(* IEC 61131-3 sources: plc-process-lib/tests/POUs/Suites/FB_Valve_Test, 85 files *)

(* ---- ActTimeAccumulatesInRetain.method.decl.st ---- *)
// Время работы привода: 12,5 с с включённым выходом — 12 с в stRetain (доля 0,5 с в накопителе), часы в
// Sts; пока стоит — не копится; шаг времени 60 с идёт в счёт не больше DT_ACCUM_MAX = 10 с. xResetMaint
// обнуляет время «с ТО», полное время не трогает.
METHOD PRIVATE ActTimeAccumulatesInRetain
VAR
    fbTime   : FB_FakeTime;       // подменное время, старт 1 ч
    fbVlv    : FB_Valve;          // арматура под тестом
    stCmd    : ST_ValveCmd;       // команды HMI
    stRetain : ST_DeviceRetain;   // режим Manual по умолчанию, счётчики
    stCfg    : ST_ValveCfg;       // конфигурация (умолчания: Motorized, ZSO и ZSC)
    iStep    : INT;               // шаг цикла
END_VAR

(* ---- ActTimeAccumulatesInRetain.method.impl.st ---- *)
coUnit.TEST('Valve_ActTime_AccumulatesInRetain');

stCfg.tTravel := T#120S;
stRetain.udiOpTime_s := 7190;
fbVlv.xZsc := TRUE;
fbVlv(itfTime := fbTime, stCmd := stCmd, stRetain := stRetain, stCfg := stCfg);
stCmd.xOpen := TRUE;
// t0: выход включён
fbVlv(itfTime := fbTime, stCmd := stCmd, stRetain := stRetain, stCfg := stCfg);
fbVlv.xZsc := FALSE;
FOR iStep := 1 TO 125 DO                                                // 12,5 с
    fbTime.Advance(tStep := T#100MS);
    fbVlv(itfTime := fbTime, stCmd := stCmd, stRetain := stRetain, stCfg := stCfg);
END_FOR
stCmd.xStop := TRUE;
// без шага времени
fbVlv(itfTime := fbTime, stCmd := stCmd, stRetain := stRetain, stCfg := stCfg);
// источник: tools/reference/valve_reference.py, сценарий valve_act_time: 12 с, в накопителе 0,5 с
AssertEquals_UDINT(Expected := 7202, Actual := stRetain.udiOpTime_s, Message := 'total run time 7190 + 12 s');
AssertEquals_UDINT(Expected := 12, Actual := stRetain.udiOpTimeMaint_s, Message := 'run time since maintenance 12 s');
// источник: tools/reference/valve_reference.py, сценарий valve_act_time: hours of 7190 + 12 s
AssertEquals_REAL(Expected := 2.0005555, Actual := fbVlv.stSts.rActTime_h, Delta := 1.0E-6,
                  Message := 'run time in hours');
FOR iStep := 1 TO 20 DO
    fbTime.Advance(tStep := T#100MS);
    fbVlv(itfTime := fbTime, stCmd := stCmd, stRetain := stRetain, stCfg := stCfg);
END_FOR
AssertEquals_UDINT(Expected := 7202, Actual := stRetain.udiOpTime_s, Message := 'no accumulation at rest');
stCmd.xOpen := TRUE;
fbVlv(itfTime := fbTime, stCmd := stCmd, stRetain := stRetain, stCfg := stCfg);
fbTime.Advance(tStep := T#1M);
// один шаг 60 с
fbVlv(itfTime := fbTime, stCmd := stCmd, stRetain := stRetain, stCfg := stCfg);
// источник: tools/reference/valve_reference.py, сценарий valve_act_time: one 60 s step = 10 s (0,5 + 10 с)
AssertEquals_UDINT(Expected := 7212, Actual := stRetain.udiOpTime_s, Message := 'large step bounded by DT_ACCUM_MAX');
stCmd.xResetMaint := TRUE;
fbVlv(itfTime := fbTime, stCmd := stCmd, stRetain := stRetain, stCfg := stCfg);
AssertEquals_UDINT(Expected := 0, Actual := stRetain.udiOpTimeMaint_s,
                   Message := 'xResetMaint clears run time since maintenance');
AssertEquals_UDINT(Expected := 7212, Actual := stRetain.udiOpTime_s, Message := 'total run time kept');

coUnit.TEST_FINISHED();

(* ---- AutoToManualBumpless.method.decl.st ---- *)
// Auto открывает; переход в Manual: цель := текущее направление — ход продолжается до ZSO (арматура не
// дёргается).
METHOD PRIVATE AutoToManualBumpless
VAR
    fbTime   : FB_FakeTime;       // подменное время, старт 1 ч
    fbVlv    : FB_Valve;          // арматура под тестом
    stCmd    : ST_ValveCmd;       // команды HMI
    stRetain : ST_DeviceRetain;   // режим Manual по умолчанию, счётчики
    stCfg    : ST_ValveCfg;       // конфигурация (умолчания: Motorized, ZSO и ZSC)
    iStep    : INT;               // шаг цикла
END_VAR

(* ---- AutoToManualBumpless.method.impl.st ---- *)
coUnit.TEST('Valve_AutoToManual_Bumpless');

stRetain.eRemoteMode := E_DeviceMode.Auto;
fbVlv.xAutoOpen := TRUE;
fbVlv.xZsc := TRUE;
fbVlv(itfTime := fbTime, stCmd := stCmd, stRetain := stRetain, stCfg := stCfg);
AssertTrue(Condition := fbVlv.stSts.eState = E_ValveState.Opening, Message := 'Auto opens on first call');
fbVlv.xZsc := FALSE;
FOR iStep := 1 TO 10 DO
    fbTime.Advance(tStep := T#100MS);
    fbVlv(itfTime := fbTime, stCmd := stCmd, stRetain := stRetain, stCfg := stCfg);
END_FOR
stCmd.stCommon.xSetManual := TRUE;
fbVlv.xAutoOpen := FALSE;
fbTime.Advance(tStep := T#100MS);
fbVlv(itfTime := fbTime, stCmd := stCmd, stRetain := stRetain, stCfg := stCfg);
AssertTrue(Condition := fbVlv.Mode = E_DeviceMode.Manual, Message := 'Manual');
AssertTrue(Condition := fbVlv.stSts.eState = E_ValveState.Opening, Message := 'keeps direction');
AssertTrue(Condition := fbVlv.xQOpen, Message := 'output kept');
FOR iStep := 1 TO 10 DO
    fbTime.Advance(tStep := T#100MS);
    fbVlv.xZso := iStep >= 10;
    fbVlv(itfTime := fbTime, stCmd := stCmd, stRetain := stRetain, stCfg := stCfg);
END_FOR
AssertTrue(Condition := fbVlv.stSts.eState = E_ValveState.Open, Message := 'Open on ZSO');
AssertFalse(Condition := fbVlv.xQOpen, Message := 'output off');

coUnit.TEST_FINISHED();

(* ---- BothLimitsSetsFailureOutputsOff.method.decl.st ---- *)
// Auto, закрыта. Залип ZSO — оба концевика: до tLimitFilter (0,5 с) состояние держится, на 0,5 с —
// BothLimits (wFault бит 2, Failure, тревога слота 2). Запрос автоматики «открыть» выходы не включает,
// Available = FALSE. Отказ не фиксируется: концевик исправен — отказ снят без Reset, Auto ведёт к цели.
METHOD PRIVATE BothLimitsSetsFailureOutputsOff
VAR
    fbTime   : FB_FakeTime;       // подменное время, старт 1 ч
    fbVlv    : FB_Valve;          // арматура под тестом
    stCmd    : ST_ValveCmd;       // команды HMI
    stRetain : ST_DeviceRetain;   // режим Manual по умолчанию, счётчики
    stCfg    : ST_ValveCfg;       // конфигурация (умолчания: Motorized, ZSO и ZSC)
    iStep    : INT;               // шаг цикла
    itfAlm   : I_Alarm;           // слот тревоги через интерфейс
END_VAR

(* ---- BothLimitsSetsFailureOutputsOff.method.impl.st ---- *)
coUnit.TEST('Valve_BothLimits_SetsFailureOutputsOff');

stRetain.eRemoteMode := E_DeviceMode.Auto;
fbVlv.xAutoOpen := FALSE;
fbVlv.xZsc := TRUE;
// Auto, закрыта
fbVlv(itfTime := fbTime, stCmd := stCmd, stRetain := stRetain, stCfg := stCfg);
AssertTrue(Condition := fbVlv.Mode = E_DeviceMode.Auto, Message := 'Auto from retain');
AssertTrue(Condition := fbVlv.stSts.eState = E_ValveState.Closed, Message := 'Closed');
fbVlv.xZso := TRUE;
// t0: оба концевика
fbVlv(itfTime := fbTime, stCmd := stCmd, stRetain := stRetain, stCfg := stCfg);
FOR iStep := 1 TO 4 DO                                                  // t0 + 0,4 с
    fbTime.Advance(tStep := T#100MS);
    fbVlv(itfTime := fbTime, stCmd := stCmd, stRetain := stRetain, stCfg := stCfg);
END_FOR
AssertEquals_WORD(Expected := 0, Actual := fbVlv.stSts.stCommon.wFault, Message := 'no fault before tLimitFilter');
AssertTrue(Condition := fbVlv.stSts.eState = E_ValveState.Closed, Message := 'state held during the filter');
fbTime.Advance(tStep := T#100MS);
// t0 + 0,5 с
fbVlv(itfTime := fbTime, stCmd := stCmd, stRetain := stRetain, stCfg := stCfg);
AssertEquals_WORD(Expected := GVL_Const.VLV_FLT_BOTH_LIMITS, Actual := fbVlv.stSts.stCommon.wFault,
                  Message := 'BothLimits after tLimitFilter');
AssertTrue(Condition := fbVlv.stSts.eState = E_ValveState.Fault, Message := 'Fault state');
AssertTrue(Condition := fbVlv.Status = E_Ne107Status.Failure, Message := 'NE 107 Failure');
itfAlm := fbVlv.GetAlarm(uiIndex := E_ValveAlarm.BothLimits);
AssertTrue(Condition := itfAlm.Active, Message := 'BothLimits alarm active');
fbVlv.xAutoOpen := TRUE;
fbTime.Advance(tStep := T#100MS);
fbVlv(itfTime := fbTime, stCmd := stCmd, stRetain := stRetain, stCfg := stCfg);
AssertFalse(Condition := fbVlv.xQOpen OR fbVlv.xQClose, Message := 'outputs off while both limit switches');
AssertFalse(Condition := fbVlv.Available, Message := 'not available');
fbVlv.xZso := FALSE;
fbTime.Advance(tStep := T#100MS);
// концевик исправен
fbVlv(itfTime := fbTime, stCmd := stCmd, stRetain := stRetain, stCfg := stCfg);
AssertEquals_WORD(Expected := 0, Actual := fbVlv.stSts.stCommon.wFault, Message := 'not latched: clears without Reset');
AssertTrue(Condition := fbVlv.stSts.eState = E_ValveState.Opening, Message := 'Auto resumes towards target');
AssertTrue(Condition := fbVlv.xQOpen, Message := 'open contactor on');

coUnit.TEST_FINISHED();

(* ---- CfgChecksSetBits.method.decl.st ---- *)
// Каждая проверка CheckConfig даёт свой бит wCfgErr: тип вне перечисления; tTravel = 0; Stay у соленоида
// и eSafePos вне перечисления; закрытие по моменту без муфты и муфта у соленоида; tReverse = 0 у
// Motorized (у соленоида допустим); tResetWindow = 0; приоритет тревоги вне перечисления.
METHOD PRIVATE CfgChecksSetBits
VAR
    fbTime   : FB_FakeTime;       // подменное время, старт 1 ч
    fbVlv    : FB_Valve;          // арматура под тестом
    stCmd    : ST_ValveCmd;       // команды HMI
    stRetain : ST_DeviceRetain;   // режим Manual по умолчанию, счётчики
    stCfg    : ST_ValveCfg;       // конфигурация (умолчания: Motorized, ZSO и ZSC)
    uBad     : U_TestValveEnum;   // значения вне строгих перечислений
    stSlot   : ST_AlarmCfg;       // копия слота тревоги
END_VAR

(* ---- CloseLimitReachedGoesClosed.method.decl.st ---- *)
// Manual, задвижка открыта (ZSO). xClose: Closing, включён только xQClose; ZSC на t0 + 3,0 с — Closed,
// выход снят, xClosed. Закрытие циклом «открыто» не считается.
METHOD PRIVATE CloseLimitReachedGoesClosed
VAR
    fbTime   : FB_FakeTime;       // подменное время, старт 1 ч
    fbVlv    : FB_Valve;          // арматура под тестом
    stCmd    : ST_ValveCmd;       // команды HMI
    stRetain : ST_DeviceRetain;   // режим Manual по умолчанию, счётчики
    stCfg    : ST_ValveCfg;       // конфигурация (умолчания: Motorized, ZSO и ZSC)
    iStep    : INT;               // шаг цикла
END_VAR

(* ---- CloseLimitReachedGoesClosed.method.impl.st ---- *)
coUnit.TEST('Valve_Close_LimitReached_GoesClosed');

stCfg.tTravel := T#10S;
fbVlv.xZso := TRUE;
// t0: открыта
fbVlv(itfTime := fbTime, stCmd := stCmd, stRetain := stRetain, stCfg := stCfg);
AssertTrue(Condition := fbVlv.stSts.eState = E_ValveState.Open, Message := 'starts Open on ZSO');
stCmd.xClose := TRUE;
// t0: команда «закрыть»
fbVlv(itfTime := fbTime, stCmd := stCmd, stRetain := stRetain, stCfg := stCfg);
AssertTrue(Condition := fbVlv.stSts.eState = E_ValveState.Closing, Message := 'Closing after xClose');
AssertTrue(Condition := fbVlv.xQClose, Message := 'close contactor on');
AssertFalse(Condition := fbVlv.xQOpen, Message := 'open contactor off');
AssertFalse(Condition := stCmd.xClose, Message := 'xClose cleared');
AssertEquals_WORD(Expected := GVL_Const.VLV_STS_CLOSING,
                  Actual := fbVlv.stSts.stCommon.wStatus AND GVL_Const.VLV_STS_CLOSING, Message := 'CLOSING bit');
FOR iStep := 1 TO 29 DO                                                 // t0 + 0,1 … 2,9 с; ZSO пропал на 0,3 с
    fbTime.Advance(tStep := T#100MS);
    fbVlv.xZso := iStep < 3;
    fbVlv(itfTime := fbTime, stCmd := stCmd, stRetain := stRetain, stCfg := stCfg);
END_FOR
AssertTrue(Condition := fbVlv.xQClose, Message := 'still closing at t0 + 2.9 s');
fbTime.Advance(tStep := T#100MS);
fbVlv.xZsc := TRUE;
// t0 + 3,0 с: ZSC
fbVlv(itfTime := fbTime, stCmd := stCmd, stRetain := stRetain, stCfg := stCfg);
AssertTrue(Condition := fbVlv.stSts.eState = E_ValveState.Closed, Message := 'Closed on ZSC');
AssertFalse(Condition := fbVlv.xQClose, Message := 'contactor off at ZSC');
AssertTrue(Condition := fbVlv.xClosed, Message := 'xClosed');
AssertFalse(Condition := fbVlv.xOpened, Message := 'not xOpened');
AssertEquals_WORD(Expected := GVL_Const.VLV_STS_CLOSED,
                  Actual := fbVlv.stSts.stCommon.wStatus AND (GVL_Const.VLV_STS_OPENED OR GVL_Const.VLV_STS_CLOSED),
                  Message := 'CLOSED bit');
AssertEquals_UDINT(Expected := 0, Actual := stRetain.udiOpCount, Message := 'closing is not an open cycle');

coUnit.TEST_FINISHED();

(* ---- CloseOnTorqueCompletesClosing.method.decl.st ---- *)
// Клиновая задвижка: муфта подключена, закрытие «по моменту». Через 3 с хода сработал ZSC (стоит чуть
// раньше посадки клина) — выход держится; через 0,2 с клин сел, сработала муфта закрытия — Closed без
// отказа, выход снят, xClosed; предупреждения «положение по времени» нет. Муфта отпустила, ZSC держится —
// задвижка остаётся Closed без отказа. Муфта раньше ZSC — тест
// Valve_CloseOnTorque_TorqueBeforeZsc_LatchesTorqueTrip.
METHOD PRIVATE CloseOnTorqueCompletesClosing
VAR
    fbTime   : FB_FakeTime;       // подменное время, старт 1 ч
    fbVlv    : FB_Valve;          // арматура под тестом
    stCmd    : ST_ValveCmd;       // команды HMI
    stRetain : ST_DeviceRetain;   // режим Manual по умолчанию, счётчики
    stCfg    : ST_ValveCfg;       // конфигурация (умолчания: Motorized, ZSO и ZSC)
    iStep    : INT;               // шаг цикла
END_VAR

(* ---- CloseOnTorqueCompletesClosing.method.impl.st ---- *)
coUnit.TEST('Valve_CloseOnTorque_CompletesClosing');

stCfg.xTorqueUsed := TRUE;
stCfg.xCloseOnTorque := TRUE;
fbVlv.xZso := TRUE;
fbVlv(itfTime := fbTime, stCmd := stCmd, stRetain := stRetain, stCfg := stCfg);
stCmd.xClose := TRUE;
fbVlv(itfTime := fbTime, stCmd := stCmd, stRetain := stRetain, stCfg := stCfg);
fbVlv.xZso := FALSE;
FOR iStep := 1 TO 30 DO                                                 // закрывается 3 с
    fbTime.Advance(tStep := T#100MS);
    fbVlv(itfTime := fbTime, stCmd := stCmd, stRetain := stRetain, stCfg := stCfg);
END_FOR
fbVlv.xZsc := TRUE;
FOR iStep := 1 TO 2 DO                                                  // ZSC: клин дожимается 0,2 с
    fbTime.Advance(tStep := T#100MS);
    fbVlv(itfTime := fbTime, stCmd := stCmd, stRetain := stRetain, stCfg := stCfg);
END_FOR
AssertTrue(Condition := fbVlv.xQClose, Message := 'output held on ZSC until torque');
fbVlv.xTorqueClose := TRUE;
fbTime.Advance(tStep := T#100MS);
// клин сел: муфта закрытия
fbVlv(itfTime := fbTime, stCmd := stCmd, stRetain := stRetain, stCfg := stCfg);
AssertTrue(Condition := fbVlv.stSts.eState = E_ValveState.Closed, Message := 'Closed on torque');
AssertFalse(Condition := fbVlv.xQClose, Message := 'output off');
AssertEquals_WORD(Expected := 0, Actual := fbVlv.stSts.stCommon.wFault, Message := 'no torque trip');
AssertTrue(Condition := fbVlv.xClosed, Message := 'xClosed');
AssertEquals_WORD(Expected := 0, Actual := fbVlv.stSts.stCommon.wWarning AND GVL_Const.VLV_WRN_POSITION_BY_TIME,
                  Message := 'closed by torque, not by time');
fbVlv.xTorqueClose := FALSE;
FOR iStep := 1 TO 20 DO                                                 // 2 с: муфта отпустила, ZSC держится
    fbTime.Advance(tStep := T#100MS);
    fbVlv(itfTime := fbTime, stCmd := stCmd, stRetain := stRetain, stCfg := stCfg);
END_FOR
AssertEquals_WORD(Expected := 0, Actual := fbVlv.stSts.stCommon.wFault, Message := 'no fault after torque released');
AssertTrue(Condition := fbVlv.stSts.eState = E_ValveState.Closed, Message := 'stays Closed');

coUnit.TEST_FINISHED();

(* ---- CloseOnTorqueNoZscTorqueMissingSetsFailToClose.method.decl.st ---- *)
// Клиновая задвижка без ZSC (xZscUsed = FALSE), закрытие «по моменту», tTravel = 10 с. Муфта закрытия
// так и не сработала: на t0 + 9,9 с ещё Closing и выход «закрывать» держится, ровно на t0 + 10,0 с —
// FailToClose, выход снят, xClosed нет. Положения «закрыто по времени» у закрытия по моменту нет: его
// подтверждает только муфта.
METHOD PRIVATE CloseOnTorqueNoZscTorqueMissingSetsFailToClose
VAR
    fbTime   : FB_FakeTime;       // подменное время, старт 1 ч
    fbVlv    : FB_Valve;          // арматура под тестом
    stCmd    : ST_ValveCmd;       // команды HMI
    stRetain : ST_DeviceRetain;   // режим Manual по умолчанию, счётчики
    stCfg    : ST_ValveCfg;       // конфигурация: без ZSC, закрытие по моменту
    iStep    : INT;               // шаг цикла
END_VAR

(* ---- CloseOnTorqueNoZscTorqueMissingSetsFailToClose.method.impl.st ---- *)
coUnit.TEST('Valve_CloseOnTorqueNoZsc_TorqueMissing_SetsFailToClose');

stCfg.xZscUsed := FALSE;
stCfg.xTorqueUsed := TRUE;
stCfg.xCloseOnTorque := TRUE;
stCfg.tTravel := T#10S;
fbVlv.xZso := TRUE;
fbVlv(itfTime := fbTime, stCmd := stCmd, stRetain := stRetain, stCfg := stCfg);
stCmd.xClose := TRUE;
// t0: Closing
fbVlv(itfTime := fbTime, stCmd := stCmd, stRetain := stRetain, stCfg := stCfg);
fbVlv.xZso := FALSE;
FOR iStep := 1 TO 99 DO                                                 // до t0 + 9,9 с, муфты нет
    fbTime.Advance(tStep := T#100MS);
    fbVlv(itfTime := fbTime, stCmd := stCmd, stRetain := stRetain, stCfg := stCfg);
END_FOR
AssertTrue(Condition := fbVlv.stSts.eState = E_ValveState.Closing, Message := 'still closing at t0 + 9.9 s');
AssertTrue(Condition := fbVlv.xQClose, Message := 'close output held until torque');
fbTime.Advance(tStep := T#100MS);
// t0 + 10,0 с
fbVlv(itfTime := fbTime, stCmd := stCmd, stRetain := stRetain, stCfg := stCfg);
AssertTrue(Condition := fbVlv.stSts.eState = E_ValveState.Fault, Message := 'Fault at tTravel, not closed by time');
AssertEquals_WORD(Expected := GVL_Const.VLV_FLT_FAIL_TO_CLOSE, Actual := fbVlv.stSts.stCommon.wFault,
                  Message := 'wFault FailToClose');
AssertFalse(Condition := fbVlv.xQClose, Message := 'output off on timeout');
AssertFalse(Condition := fbVlv.xClosed, Message := 'not reported closed');

coUnit.TEST_FINISHED();

(* ---- CloseOnTorqueTorqueBeforeZscLatchesTorqueTrip.method.decl.st ---- *)
// Клиновая задвижка, закрытие «по моменту», ZSC подключён. Муфта закрытия сработала на t0 + 3 с, а
// ZSC — нет: ZSC настроен чуть раньше посадки клина (VLV-19), значит, это не посадка, а заклинивание или
// посторонний предмет — TorqueTrip, выход снят, xClosed нет. Тот же ход без ZSC (xZscUsed = FALSE):
// муфта — штатное окончание закрытия, Closed без отказа, и после того как муфта отпустила, задвижка
// остаётся Closed.
METHOD PRIVATE CloseOnTorqueTorqueBeforeZscLatchesTorqueTrip
VAR
    fbTime    : FB_FakeTime;       // подменное время, старт 1 ч
    fbVlv     : FB_Valve;          // задвижка с ZSC
    stCmd     : ST_ValveCmd;       // команды HMI
    stRetain  : ST_DeviceRetain;   // режим Manual по умолчанию, счётчики
    stCfg     : ST_ValveCfg;       // конфигурация (умолчания: Motorized, ZSO и ZSC)
    fbVlv2    : FB_Valve;          // задвижка без ZSC
    stCmd2    : ST_ValveCmd;       // команды HMI второй задвижки
    stRetain2 : ST_DeviceRetain;   // режим Manual по умолчанию
    stCfg2    : ST_ValveCfg;       // конфигурация второй задвижки
    iStep     : INT;               // шаг цикла
END_VAR

(* ---- CloseOnTorqueTorqueBeforeZscLatchesTorqueTrip.method.impl.st ---- *)
coUnit.TEST('Valve_CloseOnTorque_TorqueBeforeZsc_LatchesTorqueTrip');

stCfg.xTorqueUsed := TRUE;
stCfg.xCloseOnTorque := TRUE;
fbVlv.xZso := TRUE;
fbVlv(itfTime := fbTime, stCmd := stCmd, stRetain := stRetain, stCfg := stCfg);
stCmd.xClose := TRUE;
fbVlv(itfTime := fbTime, stCmd := stCmd, stRetain := stRetain, stCfg := stCfg);
fbVlv.xZso := FALSE;
FOR iStep := 1 TO 30 DO                                                 // закрывается 3 с
    fbTime.Advance(tStep := T#100MS);
    fbVlv(itfTime := fbTime, stCmd := stCmd, stRetain := stRetain, stCfg := stCfg);
END_FOR
fbVlv.xTorqueClose := TRUE;
fbTime.Advance(tStep := T#100MS);
// муфта раньше ZSC
fbVlv(itfTime := fbTime, stCmd := stCmd, stRetain := stRetain, stCfg := stCfg);
AssertTrue(Condition := fbVlv.stSts.eState = E_ValveState.Fault, Message := 'torque before ZSC: Fault');
AssertEquals_WORD(Expected := GVL_Const.VLV_FLT_TORQUE_TRIP, Actual := fbVlv.stSts.stCommon.wFault,
                  Message := 'wFault TorqueTrip');
AssertFalse(Condition := fbVlv.xQClose, Message := 'output off');
AssertFalse(Condition := fbVlv.xClosed, Message := 'not reported closed');

stCfg2.xZscUsed := FALSE;
stCfg2.xTorqueUsed := TRUE;
stCfg2.xCloseOnTorque := TRUE;
fbVlv2.xZso := TRUE;
fbVlv2(itfTime := fbTime, stCmd := stCmd2, stRetain := stRetain2, stCfg := stCfg2);
stCmd2.xClose := TRUE;
fbVlv2(itfTime := fbTime, stCmd := stCmd2, stRetain := stRetain2, stCfg := stCfg2);
fbVlv2.xZso := FALSE;
FOR iStep := 1 TO 30 DO                                                 // закрывается 3 с
    fbTime.Advance(tStep := T#100MS);
    fbVlv2(itfTime := fbTime, stCmd := stCmd2, stRetain := stRetain2, stCfg := stCfg2);
END_FOR
fbVlv2.xTorqueClose := TRUE;
fbTime.Advance(tStep := T#100MS);
// без ZSC муфта — окончание закрытия
fbVlv2(itfTime := fbTime, stCmd := stCmd2, stRetain := stRetain2, stCfg := stCfg2);
AssertTrue(Condition := fbVlv2.stSts.eState = E_ValveState.Closed, Message := 'no ZSC: Closed on torque');
AssertEquals_WORD(Expected := 0, Actual := fbVlv2.stSts.stCommon.wFault, Message := 'no ZSC: no torque trip');
AssertFalse(Condition := fbVlv2.xQClose, Message := 'no ZSC: output off');
AssertTrue(Condition := fbVlv2.xClosed, Message := 'no ZSC: xClosed');
fbVlv2.xTorqueClose := FALSE;
FOR iStep := 1 TO 20 DO                                                 // муфта отпустила, 2 с
    fbTime.Advance(tStep := T#100MS);
    fbVlv2(itfTime := fbTime, stCmd := stCmd2, stRetain := stRetain2, stCfg := stCfg2);
END_FOR
AssertTrue(Condition := fbVlv2.stSts.eState = E_ValveState.Closed, Message := 'no ZSC: stays Closed');
AssertEquals_WORD(Expected := 0, Actual := fbVlv2.stSts.stCommon.wFault, Message := 'no ZSC: still no fault');

coUnit.TEST_FINISHED();

(* ---- CloseOnTorqueZscAloneKeepsDrivingUntilTimeout.method.decl.st ---- *)
// Клиновая задвижка, закрытие «по моменту», tTravel = 10 с. ZSC сработал на t0 + 3 с (концевик стоит
// чуть раньше посадки клина): выход «закрывать» не снимается — клин дожимается до муфты, xClosed нет.
// Муфта так и не сработала: ровно на t0 + 10,0 с — FailToClose, выход снят; положение по ZSC видно в
// xClosed. Reset снимает отказ — далее состояние по концевикам (Closed).
METHOD PRIVATE CloseOnTorqueZscAloneKeepsDrivingUntilTimeout
VAR
    fbTime   : FB_FakeTime;       // подменное время, старт 1 ч
    fbVlv    : FB_Valve;          // арматура под тестом
    stCmd    : ST_ValveCmd;       // команды HMI
    stRetain : ST_DeviceRetain;   // режим Manual по умолчанию, счётчики
    stCfg    : ST_ValveCfg;       // конфигурация (умолчания: Motorized, ZSO и ZSC)
    iStep    : INT;               // шаг цикла
END_VAR

(* ---- CloseOnTorqueZscAloneKeepsDrivingUntilTimeout.method.impl.st ---- *)
coUnit.TEST('Valve_CloseOnTorque_ZscAloneKeepsDrivingUntilTimeout');

stCfg.tTravel := T#10S;
stCfg.xTorqueUsed := TRUE;
stCfg.xCloseOnTorque := TRUE;
fbVlv.xZso := TRUE;
// t0: открыта
fbVlv(itfTime := fbTime, stCmd := stCmd, stRetain := stRetain, stCfg := stCfg);
stCmd.xClose := TRUE;
// t0: Closing
fbVlv(itfTime := fbTime, stCmd := stCmd, stRetain := stRetain, stCfg := stCfg);
fbVlv.xZso := FALSE;
FOR iStep := 1 TO 30 DO                                                 // до t0 + 3,0 с
    fbTime.Advance(tStep := T#100MS);
    fbVlv(itfTime := fbTime, stCmd := stCmd, stRetain := stRetain, stCfg := stCfg);
END_FOR
fbVlv.xZsc := TRUE;
FOR iStep := 1 TO 69 DO                                                 // ZSC есть, муфты нет: до t0 + 9,9 с
    fbTime.Advance(tStep := T#100MS);
    fbVlv(itfTime := fbTime, stCmd := stCmd, stRetain := stRetain, stCfg := stCfg);
END_FOR
AssertTrue(Condition := fbVlv.stSts.eState = E_ValveState.Closing, Message := 'still closing on ZSC alone');
AssertTrue(Condition := fbVlv.xQClose, Message := 'close output held until torque');
AssertFalse(Condition := fbVlv.xClosed, Message := 'not closed before torque');
AssertEquals_WORD(Expected := 0, Actual := fbVlv.stSts.stCommon.wFault, Message := 'no fault before tTravel');
fbTime.Advance(tStep := T#100MS);
// t0 + 10,0 с: муфта не сработала
fbVlv(itfTime := fbTime, stCmd := stCmd, stRetain := stRetain, stCfg := stCfg);
AssertTrue(Condition := fbVlv.stSts.eState = E_ValveState.Fault, Message := 'Fault at tTravel');
AssertEquals_WORD(Expected := GVL_Const.VLV_FLT_FAIL_TO_CLOSE, Actual := fbVlv.stSts.stCommon.wFault,
                  Message := 'wFault FailToClose');
AssertFalse(Condition := fbVlv.xQClose, Message := 'output off on timeout');
AssertTrue(Condition := fbVlv.xClosed, Message := 'ZSC position visible in Fault');
stCmd.stCommon.xReset := TRUE;
fbVlv(itfTime := fbTime, stCmd := stCmd, stRetain := stRetain, stCfg := stCfg);
AssertEquals_WORD(Expected := 0, Actual := fbVlv.stSts.stCommon.wFault, Message := 'cleared by Reset');
AssertTrue(Condition := fbVlv.stSts.eState = E_ValveState.Closed, Message := 'Closed by ZSC after Reset');
AssertFalse(Condition := fbVlv.xQClose, Message := 'no output after Reset');

coUnit.TEST_FINISHED();

(* ---- CyclesCountedOnOpen.method.decl.st ---- *)
// Цикл — вход в Open, если прошлое крайнее положение не Open: открыть (1), закрыть (1), открыть (2) —
// stRetain и stSts. Неполный ход Open -> стоп -> снова Open циклом не считается. xResetMaint обнуляет
// счётчик «с ТО», полный не трогает. Перед каждой сменой направления арматура стоит 1 с: встречный ход
// начинается не раньше tReverse после снятия выхода (тест Valve_ReverseAfterEndStop_WaitsReversePause).
METHOD PRIVATE CyclesCountedOnOpen
VAR
    fbTime   : FB_FakeTime;       // подменное время, старт 1 ч
    fbVlv    : FB_Valve;          // арматура под тестом
    stCmd    : ST_ValveCmd;       // команды HMI
    stRetain : ST_DeviceRetain;   // режим Manual по умолчанию, счётчики
    stCfg    : ST_ValveCfg;       // конфигурация (умолчания: Motorized, ZSO и ZSC)
    iStep    : INT;               // шаг цикла
END_VAR

(* ---- CyclesCountedOnOpen.method.impl.st ---- *)
coUnit.TEST('Valve_Cycles_CountedOnOpen');

fbVlv.xZsc := TRUE;
fbVlv(itfTime := fbTime, stCmd := stCmd, stRetain := stRetain, stCfg := stCfg);
stCmd.xOpen := TRUE;
fbVlv(itfTime := fbTime, stCmd := stCmd, stRetain := stRetain, stCfg := stCfg);
FOR iStep := 1 TO 10 DO
    fbTime.Advance(tStep := T#100MS);
    fbVlv.xZsc := FALSE;
    fbVlv.xZso := iStep >= 10;
    fbVlv(itfTime := fbTime, stCmd := stCmd, stRetain := stRetain, stCfg := stCfg);
END_FOR
AssertEquals_UDINT(Expected := 1, Actual := stRetain.udiOpCount, Message := 'first open: 1');
FOR iStep := 1 TO 10 DO                                                 // стоит 1 с (выбег, tReverse)
    fbTime.Advance(tStep := T#100MS);
    fbVlv(itfTime := fbTime, stCmd := stCmd, stRetain := stRetain, stCfg := stCfg);
END_FOR
stCmd.xClose := TRUE;
fbVlv(itfTime := fbTime, stCmd := stCmd, stRetain := stRetain, stCfg := stCfg);
FOR iStep := 1 TO 10 DO
    fbTime.Advance(tStep := T#100MS);
    fbVlv.xZso := FALSE;
    fbVlv.xZsc := iStep >= 10;
    fbVlv(itfTime := fbTime, stCmd := stCmd, stRetain := stRetain, stCfg := stCfg);
END_FOR
AssertTrue(Condition := fbVlv.stSts.eState = E_ValveState.Closed, Message := 'Closed');
AssertEquals_UDINT(Expected := 1, Actual := stRetain.udiOpCount, Message := 'closing does not count');
FOR iStep := 1 TO 10 DO                                                 // стоит 1 с (выбег, tReverse)
    fbTime.Advance(tStep := T#100MS);
    fbVlv(itfTime := fbTime, stCmd := stCmd, stRetain := stRetain, stCfg := stCfg);
END_FOR
stCmd.xOpen := TRUE;
fbVlv(itfTime := fbTime, stCmd := stCmd, stRetain := stRetain, stCfg := stCfg);
FOR iStep := 1 TO 10 DO
    fbTime.Advance(tStep := T#100MS);
    fbVlv.xZsc := FALSE;
    fbVlv.xZso := iStep >= 10;
    fbVlv(itfTime := fbTime, stCmd := stCmd, stRetain := stRetain, stCfg := stCfg);
END_FOR
AssertEquals_UDINT(Expected := 2, Actual := stRetain.udiOpCount, Message := 'second open: 2');
AssertEquals_UDINT(Expected := 2, Actual := stRetain.udiOpCountMaint, Message := 'maintenance counter 2');
AssertEquals_UDINT(Expected := 2, Actual := fbVlv.stSts.udiCycles, Message := 'Sts udiCycles');
AssertEquals_UDINT(Expected := 2, Actual := fbVlv.stSts.udiCyclesMaint, Message := 'Sts udiCyclesMaint');
FOR iStep := 1 TO 10 DO                                                 // стоит 1 с (выбег, tReverse)
    fbTime.Advance(tStep := T#100MS);
    fbVlv(itfTime := fbTime, stCmd := stCmd, stRetain := stRetain, stCfg := stCfg);
END_FOR
stCmd.xClose := TRUE;
fbVlv(itfTime := fbTime, stCmd := stCmd, stRetain := stRetain, stCfg := stCfg);
FOR iStep := 1 TO 5 DO
    fbTime.Advance(tStep := T#100MS);
    fbVlv.xZso := FALSE;
    fbVlv(itfTime := fbTime, stCmd := stCmd, stRetain := stRetain, stCfg := stCfg);
END_FOR
stCmd.xStop := TRUE;
fbVlv(itfTime := fbTime, stCmd := stCmd, stRetain := stRetain, stCfg := stCfg);
FOR iStep := 1 TO 10 DO                                                 // стоит 1 с (выбег, tReverse)
    fbTime.Advance(tStep := T#100MS);
    fbVlv(itfTime := fbTime, stCmd := stCmd, stRetain := stRetain, stCfg := stCfg);
END_FOR
stCmd.xOpen := TRUE;
fbVlv(itfTime := fbTime, stCmd := stCmd, stRetain := stRetain, stCfg := stCfg);
FOR iStep := 1 TO 5 DO
    fbTime.Advance(tStep := T#100MS);
    fbVlv.xZso := iStep >= 5;
    fbVlv(itfTime := fbTime, stCmd := stCmd, stRetain := stRetain, stCfg := stCfg);
END_FOR
AssertTrue(Condition := fbVlv.stSts.eState = E_ValveState.Open, Message := 'Open again');
AssertEquals_UDINT(Expected := 2, Actual := stRetain.udiOpCount,
                   Message := 'partial stroke back to Open is not a cycle');
stCmd.xResetMaint := TRUE;
fbVlv(itfTime := fbTime, stCmd := stCmd, stRetain := stRetain, stCfg := stCfg);
AssertEquals_UDINT(Expected := 0, Actual := stRetain.udiOpCountMaint, Message := 'maintenance counter reset');
AssertEquals_UDINT(Expected := 2, Actual := stRetain.udiOpCount, Message := 'total kept');
AssertTrue(Condition := fbVlv.stSts.stCommon.eCmdResult = E_CmdResult.Accepted, Message := 'xResetMaint accepted');
AssertFalse(Condition := stCmd.xResetMaint, Message := 'xResetMaint cleared');

coUnit.TEST_FINISHED();

(* ---- DefaultCfgPassesCheck.method.decl.st ---- *)
// Умолчания ST_ValveCfg проходят CheckConfig; тип в stCommon — Valve, слотов тревог 7; приоритеты по
// умолчанию (FailToOpen — Medium, InterlockAct — None); слот 7 не используется; NE 107 Good.
METHOD PRIVATE DefaultCfgPassesCheck
VAR
    fbTime   : FB_FakeTime;       // подменное время, старт 1 ч
    fbVlv    : FB_Valve;          // арматура под тестом
    stCmd    : ST_ValveCmd;       // команды HMI
    stRetain : ST_DeviceRetain;   // режим Manual по умолчанию, счётчики
    stCfg    : ST_ValveCfg;       // конфигурация (умолчания: Motorized, ZSO и ZSC)
    itfAlm   : I_Alarm;           // слот тревоги через интерфейс
END_VAR

(* ---- ExtFaultTripsAndResetRejectedWhileActive.method.decl.st ---- *)
// Внешняя авария в ходе: Fault, выход снят, тревога слота 5 с номером udiAlarmIdBase + 5. Reset при
// действующей причине: Accepted сразу, окно tResetWindow = 3 с; до конца окна второго результата нет,
// ровно на 3 с — RejectedFault, отказ остаётся. Причина ушла — отказ держится до Reset; Reset снимает.
METHOD PRIVATE ExtFaultTripsAndResetRejectedWhileActive
VAR
    fbTime   : FB_FakeTime;       // подменное время, старт 1 ч
    fbVlv    : FB_Valve;          // арматура под тестом
    stCmd    : ST_ValveCmd;       // команды HMI
    stRetain : ST_DeviceRetain;   // режим Manual по умолчанию, счётчики
    stCfg    : ST_ValveCfg;       // конфигурация (умолчания: Motorized, ZSO и ZSC)
    iStep    : INT;               // шаг цикла
    itfAlm   : I_Alarm;           // слот тревоги через интерфейс
    uiSeq    : UINT;              // номер команды до Reset
END_VAR

(* ---- ExtFaultTripsAndResetRejectedWhileActive.method.impl.st ---- *)
coUnit.TEST('Valve_ExtFault_TripsAndResetRejectedWhileActive');

stCfg.udiAlarmIdBase := 120;
fbVlv.xZsc := TRUE;
fbVlv(itfTime := fbTime, stCmd := stCmd, stRetain := stRetain, stCfg := stCfg);
stCmd.xOpen := TRUE;
fbVlv(itfTime := fbTime, stCmd := stCmd, stRetain := stRetain, stCfg := stCfg);
fbVlv.xZsc := FALSE;
fbTime.Advance(tStep := T#100MS);
fbVlv(itfTime := fbTime, stCmd := stCmd, stRetain := stRetain, stCfg := stCfg);
fbVlv.xExtFault := TRUE;
fbTime.Advance(tStep := T#100MS);
fbVlv(itfTime := fbTime, stCmd := stCmd, stRetain := stRetain, stCfg := stCfg);
AssertTrue(Condition := fbVlv.stSts.eState = E_ValveState.Fault, Message := 'Fault on external fault');
AssertFalse(Condition := fbVlv.xQOpen, Message := 'output off');
AssertEquals_WORD(Expected := GVL_Const.VLV_FLT_EXT_FAULT, Actual := fbVlv.stSts.stCommon.wFault,
                  Message := 'wFault ExtFault');
itfAlm := fbVlv.GetAlarm(uiIndex := E_ValveAlarm.ExtFault);
AssertEquals_UDINT(Expected := 125, Actual := itfAlm.Id, Message := 'alarm id = base + slot');
AssertTrue(Condition := itfAlm.State = E_AlarmState.ActiveUnack, Message := 'ExtFault alarm');
uiSeq := fbVlv.stSts.stCommon.uiCmdSeq;
stCmd.stCommon.xReset := TRUE;
// t1: Reset, причина действует
fbVlv(itfTime := fbTime, stCmd := stCmd, stRetain := stRetain, stCfg := stCfg);
AssertTrue(Condition := fbVlv.stSts.stCommon.eCmdResult = E_CmdResult.Accepted, Message := 'Reset accepted');
AssertEquals_UINT(Expected := uiSeq + 1, Actual := fbVlv.stSts.stCommon.uiCmdSeq, Message := 'one result so far');
FOR iStep := 1 TO 29 DO                                                 // t1 + 2,9 с
    fbTime.Advance(tStep := T#100MS);
    fbVlv(itfTime := fbTime, stCmd := stCmd, stRetain := stRetain, stCfg := stCfg);
END_FOR
AssertEquals_UINT(Expected := uiSeq + 1, Actual := fbVlv.stSts.stCommon.uiCmdSeq,
                  Message := 'no second result before the window ends');
fbTime.Advance(tStep := T#100MS);
// t1 + 3,0 с
fbVlv(itfTime := fbTime, stCmd := stCmd, stRetain := stRetain, stCfg := stCfg);
AssertTrue(Condition := fbVlv.stSts.stCommon.eCmdResult = E_CmdResult.RejectedFault,
           Message := 'RejectedFault at the window end');
AssertEquals_UINT(Expected := uiSeq + 2, Actual := fbVlv.stSts.stCommon.uiCmdSeq, Message := 'second result');
AssertEquals_WORD(Expected := GVL_Const.VLV_FLT_EXT_FAULT, Actual := fbVlv.stSts.stCommon.wFault,
                  Message := 'still faulted');
fbVlv.xExtFault := FALSE;
fbTime.Advance(tStep := T#100MS);
fbVlv(itfTime := fbTime, stCmd := stCmd, stRetain := stRetain, stCfg := stCfg);
AssertEquals_WORD(Expected := GVL_Const.VLV_FLT_EXT_FAULT, Actual := fbVlv.stSts.stCommon.wFault,
                  Message := 'latched after the cause is gone');
stCmd.stCommon.xReset := TRUE;
fbVlv(itfTime := fbTime, stCmd := stCmd, stRetain := stRetain, stCfg := stCfg);
AssertEquals_WORD(Expected := 0, Actual := fbVlv.stSts.stCommon.wFault, Message := 'cleared by Reset');
AssertTrue(Condition := fbVlv.stSts.stCommon.eCmdResult = E_CmdResult.Accepted, Message := 'Reset accepted');
fbTime.Advance(tStep := T#100MS);
fbVlv(itfTime := fbTime, stCmd := stCmd, stRetain := stRetain, stCfg := stCfg);
AssertTrue(Condition := itfAlm.State = E_AlarmState.Normal, Message := 'alarm Normal after Reset');
AssertTrue(Condition := fbVlv.stSts.eState = E_ValveState.Intermediate, Message := 'Intermediate');

coUnit.TEST_FINISHED();

(* ---- InterlockAfterPositionLostDrivesSafe.method.decl.st ---- *)
// Задвижка в Auto открыта по ZSO; ZSO пропал (обрыв) — через tLimitFilter зафиксирован PositionLost, выходов нет.
// Блокировка (Closed): задвижка закрывается (VLV-20); ход заканчивается по ZSC — он согласован (ZSO нет). Отказ
// держится до Reset; после Reset — Closed по концевикам, движения нет (уже в положении безопасности).
METHOD PRIVATE InterlockAfterPositionLostDrivesSafe
VAR
    fbTime   : FB_FakeTime;       // подменное время, старт 1 ч
    fbVlv    : FB_Valve;          // арматура под тестом
    stCmd    : ST_ValveCmd;       // команды HMI
    stRetain : ST_DeviceRetain;   // режим, счётчики
    stCfg    : ST_ValveCfg;       // конфигурация (умолчания: Motorized, ZSO и ZSC)
    iStep    : INT;               // шаг цикла
END_VAR

(* ---- InterlockAfterPositionLostDrivesSafe.method.impl.st ---- *)
coUnit.TEST('Valve_InterlockAfterPositionLost_DrivesSafe');

stRetain.eRemoteMode := E_DeviceMode.Auto;
fbVlv.xAutoOpen := TRUE;
fbVlv.xZso := TRUE;
fbVlv(itfTime := fbTime, stCmd := stCmd, stRetain := stRetain, stCfg := stCfg);       // t0: Open по ZSO
fbVlv.xZso := FALSE;                                                                   // обрыв ZSO
FOR iStep := 1 TO 6 DO                                                               // фильтр 0,5 с
    fbTime.Advance(tStep := T#100MS);
    fbVlv(itfTime := fbTime, stCmd := stCmd, stRetain := stRetain, stCfg := stCfg);
END_FOR
AssertEquals_WORD(Expected := GVL_Const.VLV_FLT_POSITION_LOST, Actual := fbVlv.stSts.stCommon.wFault,
                  Message := 'precondition: PositionLost latched');
AssertFalse(Condition := fbVlv.xQOpen OR fbVlv.xQClose, Message := 'no motion with the fault alone');
fbVlv.wInterlock := 16#0001;
fbTime.Advance(tStep := T#100MS);
fbVlv(itfTime := fbTime, stCmd := stCmd, stRetain := stRetain, stCfg := stCfg);       // t1: блокировка
AssertTrue(Condition := fbVlv.xQClose, Message := 'interlock drives Closed despite PositionLost');
FOR iStep := 1 TO 30 DO
    fbTime.Advance(tStep := T#100MS);
    fbVlv(itfTime := fbTime, stCmd := stCmd, stRetain := stRetain, stCfg := stCfg);
END_FOR
AssertTrue(Condition := fbVlv.xQClose, Message := 'still closing before ZSC');
fbVlv.xZsc := TRUE;
fbTime.Advance(tStep := T#100MS);
fbVlv(itfTime := fbTime, stCmd := stCmd, stRetain := stRetain, stCfg := stCfg);       // ZSC
AssertFalse(Condition := fbVlv.xQClose, Message := 'safe move ends on a consistent ZSC');
AssertTrue(Condition := fbVlv.xClosed, Message := 'position Closed shown');
AssertEquals_WORD(Expected := GVL_Const.VLV_FLT_POSITION_LOST, Actual := fbVlv.stSts.stCommon.wFault,
                  Message := 'fault latched until Reset');
stCmd.stCommon.xReset := TRUE;
fbTime.Advance(tStep := T#100MS);
fbVlv(itfTime := fbTime, stCmd := stCmd, stRetain := stRetain, stCfg := stCfg);
AssertEquals_WORD(Expected := 0, Actual := fbVlv.stSts.stCommon.wFault, Message := 'cleared by Reset');
AssertTrue(Condition := fbVlv.stSts.eState = E_ValveState.Closed, Message := 'Closed after Reset');
AssertFalse(Condition := fbVlv.xQOpen OR fbVlv.xQClose, Message := 'no motion: already in the safe position');

coUnit.TEST_FINISHED();

(* ---- InterlockDrivesToSafePosition.method.decl.st ---- *)
// Manual, открыта, разрешения на закрытие нет (xClose — RejectedPermit). Блокировка (биты 3 и 4) ведёт в
// положение безопасности Closed без разрешения: Closing, бит INTERLOCKED, wInterlock, первопричина —
// младший бит 3. Команды — RejectedInterlock; новый бит первопричину не меняет. После снятия блокировки
// Manual остаётся закрытым; первопричина держится до Reset.
METHOD PRIVATE InterlockDrivesToSafePosition
VAR
    fbTime   : FB_FakeTime;       // подменное время, старт 1 ч
    fbVlv    : FB_Valve;          // арматура под тестом
    stCmd    : ST_ValveCmd;       // команды HMI
    stRetain : ST_DeviceRetain;   // режим Manual по умолчанию, счётчики
    stCfg    : ST_ValveCfg;       // конфигурация (умолчания: Motorized, ZSO и ZSC)
    iStep    : INT;               // шаг цикла
END_VAR

(* ---- InterlockDrivesToSafePosition.method.impl.st ---- *)
coUnit.TEST('Valve_Interlock_DrivesToSafePosition');

fbVlv.xZso := TRUE;
fbVlv.wPermitClose := 16#0000;
// открыта, закрывать нельзя
fbVlv(itfTime := fbTime, stCmd := stCmd, stRetain := stRetain, stCfg := stCfg);
stCmd.xClose := TRUE;
fbVlv(itfTime := fbTime, stCmd := stCmd, stRetain := stRetain, stCfg := stCfg);
AssertTrue(Condition := fbVlv.stSts.stCommon.eCmdResult = E_CmdResult.RejectedPermit,
           Message := 'close without permit rejected');
AssertTrue(Condition := fbVlv.stSts.eState = E_ValveState.Open, Message := 'still Open');
fbVlv.wInterlock := 16#0018;
fbTime.Advance(tStep := T#100MS);
// блокировка
fbVlv(itfTime := fbTime, stCmd := stCmd, stRetain := stRetain, stCfg := stCfg);
AssertTrue(Condition := fbVlv.stSts.eState = E_ValveState.Closing, Message := 'interlock drives Closed');
AssertTrue(Condition := fbVlv.xQClose, Message := 'close contactor on without permit');
AssertEquals_WORD(Expected := GVL_Const.VLV_STS_INTERLOCKED,
                  Actual := fbVlv.stSts.stCommon.wStatus AND GVL_Const.VLV_STS_INTERLOCKED,
Message := 'INTERLOCKED bit');
AssertEquals_WORD(Expected := 16#0018, Actual := fbVlv.stSts.wInterlock, Message := 'active interlocks');
AssertEquals_UINT(Expected := 3, Actual := fbVlv.stSts.uiFirstOut, Message := 'first out = lowest new bit');
AssertEquals_WORD(Expected := 0, Actual := fbVlv.stSts.wPermitMissing, Message := 'no permit needed');
stCmd.xOpen := TRUE;
fbVlv.wInterlock := 16#001A;
fbTime.Advance(tStep := T#100MS);
fbVlv(itfTime := fbTime, stCmd := stCmd, stRetain := stRetain, stCfg := stCfg);
AssertTrue(Condition := fbVlv.stSts.stCommon.eCmdResult = E_CmdResult.RejectedInterlock,
           Message := 'command rejected under interlock');
AssertEquals_UINT(Expected := 3, Actual := fbVlv.stSts.uiFirstOut, Message := 'first out kept');
FOR iStep := 1 TO 10 DO
    fbTime.Advance(tStep := T#100MS);
    fbVlv.xZso := FALSE;
    fbVlv.xZsc := iStep >= 10;
    fbVlv(itfTime := fbTime, stCmd := stCmd, stRetain := stRetain, stCfg := stCfg);
END_FOR
AssertTrue(Condition := fbVlv.stSts.eState = E_ValveState.Closed, Message := 'Closed (safe position)');
fbVlv.wInterlock := 16#0000;
fbTime.Advance(tStep := T#100MS);
fbVlv(itfTime := fbTime, stCmd := stCmd, stRetain := stRetain, stCfg := stCfg);
AssertTrue(Condition := fbVlv.stSts.eState = E_ValveState.Closed, Message := 'stays Closed after the interlock');
AssertFalse(Condition := fbVlv.xQOpen, Message := 'no automatic return in Manual');
AssertEquals_UINT(Expected := 3, Actual := fbVlv.stSts.uiFirstOut, Message := 'first out held until Reset');
stCmd.stCommon.xReset := TRUE;
fbVlv(itfTime := fbTime, stCmd := stCmd, stRetain := stRetain, stCfg := stCfg);
AssertEquals_UINT(Expected := GVL_Const.NO_FIRST_OUT, Actual := fbVlv.stSts.uiFirstOut,
                  Message := 'first out cleared by Reset');

coUnit.TEST_FINISHED();

(* ---- InterlockStayStopsMotorized.method.decl.st ---- *)
// Положение безопасности Stay: блокировка в ходе останавливает электропривод (Intermediate), выходы
// сняты, бит INTERLOCKED.
METHOD PRIVATE InterlockStayStopsMotorized
VAR
    fbTime   : FB_FakeTime;       // подменное время, старт 1 ч
    fbVlv    : FB_Valve;          // арматура под тестом
    stCmd    : ST_ValveCmd;       // команды HMI
    stRetain : ST_DeviceRetain;   // режим Manual по умолчанию, счётчики
    stCfg    : ST_ValveCfg;       // конфигурация (умолчания: Motorized, ZSO и ZSC)
    iStep    : INT;               // шаг цикла
END_VAR

(* ---- InterlockStayStopsMotorized.method.impl.st ---- *)
coUnit.TEST('Valve_InterlockStay_StopsMotorized');

stCfg.eSafePos := E_ValveSafePos.Stay;
fbVlv.xZsc := TRUE;
fbVlv(itfTime := fbTime, stCmd := stCmd, stRetain := stRetain, stCfg := stCfg);
stCmd.xOpen := TRUE;
fbVlv(itfTime := fbTime, stCmd := stCmd, stRetain := stRetain, stCfg := stCfg);
fbVlv.xZsc := FALSE;
FOR iStep := 1 TO 10 DO
    fbTime.Advance(tStep := T#100MS);
    fbVlv(itfTime := fbTime, stCmd := stCmd, stRetain := stRetain, stCfg := stCfg);
END_FOR
fbVlv.wInterlock := 16#0001;
fbTime.Advance(tStep := T#100MS);
fbVlv(itfTime := fbTime, stCmd := stCmd, stRetain := stRetain, stCfg := stCfg);
AssertTrue(Condition := fbVlv.stSts.eState = E_ValveState.Intermediate, Message := 'Stay: stopped');
AssertFalse(Condition := fbVlv.xQOpen OR fbVlv.xQClose, Message := 'outputs off');
AssertEquals_WORD(Expected := GVL_Const.VLV_STS_INTERLOCKED,
                  Actual := fbVlv.stSts.stCommon.wStatus AND GVL_Const.VLV_STS_INTERLOCKED,
Message := 'INTERLOCKED bit');
AssertEquals_UINT(Expected := 0, Actual := fbVlv.stSts.uiFirstOut, Message := 'first out bit 0');

coUnit.TEST_FINISHED();

(* ---- InterlockWithBothLimitsDrivesSafe.method.decl.st ---- *)
// Задвижка в Auto открыта по ZSO; замыкание в цепи ZSC — оба концевика дольше tLimitFilter, отказ BothLimits.
// Блокировка (положение безопасности Closed): привод исправен, отказал только контроль концевиков — задвижка
// закрывается (VLV-20), состояние Fault, биты INTERLOCKED и CLOSING. Концевикам верить нельзя, поэтому ход
// заканчивается по tTravel (60 с), а не по ZSC; дальше, пока блокировка держится, ход не повторяется; оба выхода
// никогда.
METHOD PRIVATE InterlockWithBothLimitsDrivesSafe
VAR
    fbTime   : FB_FakeTime;       // подменное время, старт 1 ч
    fbVlv    : FB_Valve;          // арматура под тестом
    stCmd    : ST_ValveCmd;       // команды HMI
    stRetain : ST_DeviceRetain;   // режим, счётчики
    stCfg    : ST_ValveCfg;       // конфигурация (умолчания: Motorized, ZSO и ZSC)
    iStep    : INT;               // шаг цикла

    xCloseOn : BOOL;              // «закрывать» включено во всех вызовах хода до 59,9 с
    xBoth    : BOOL;              // оба выхода хоть раз
END_VAR

(* ---- InterlockWithBothLimitsDrivesSafe.method.impl.st ---- *)
coUnit.TEST('Valve_InterlockWithBothLimits_DrivesSafe');

stRetain.eRemoteMode := E_DeviceMode.Auto;
fbVlv.xAutoOpen := TRUE;
fbVlv.xZso := TRUE;
fbVlv(itfTime := fbTime, stCmd := stCmd, stRetain := stRetain, stCfg := stCfg);       // t0: Open по ZSO
AssertTrue(Condition := fbVlv.stSts.eState = E_ValveState.Open, Message := 'precondition: Open');
fbVlv.xZsc := TRUE;                                                                    // замыкание в цепи ZSC
FOR iStep := 1 TO 6 DO                                                               // фильтр 0,5 с
    fbTime.Advance(tStep := T#100MS);
    fbVlv(itfTime := fbTime, stCmd := stCmd, stRetain := stRetain, stCfg := stCfg);
END_FOR
AssertEquals_WORD(Expected := GVL_Const.VLV_FLT_BOTH_LIMITS, Actual := fbVlv.stSts.stCommon.wFault,
                  Message := 'precondition: BothLimits');
AssertFalse(Condition := fbVlv.xQClose, Message := 'no motion before the interlock');
fbVlv.wInterlock := 16#0001;
fbTime.Advance(tStep := T#100MS);
fbVlv(itfTime := fbTime, stCmd := stCmd, stRetain := stRetain, stCfg := stCfg);       // t1: блокировка
AssertTrue(Condition := fbVlv.xQClose, Message := 'interlock drives to the safe position despite BothLimits');
AssertFalse(Condition := fbVlv.xQOpen, Message := 'open output off');
AssertTrue(Condition := fbVlv.stSts.eState = E_ValveState.Fault, Message := 'state stays Fault');
AssertEquals_WORD(Expected := GVL_Const.VLV_STS_INTERLOCKED OR GVL_Const.VLV_STS_CLOSING,
                  Actual := fbVlv.stSts.stCommon.wStatus
                      AND (GVL_Const.VLV_STS_INTERLOCKED OR GVL_Const.VLV_STS_CLOSING),
                  Message := 'INTERLOCKED and CLOSING bits');
xCloseOn := TRUE;
FOR iStep := 1 TO 599 DO
    fbTime.Advance(tStep := T#100MS);
    fbVlv(itfTime := fbTime, stCmd := stCmd, stRetain := stRetain, stCfg := stCfg);
    xCloseOn := xCloseOn AND fbVlv.xQClose;
    xBoth := xBoth OR (fbVlv.xQOpen AND fbVlv.xQClose);
END_FOR
AssertTrue(Condition := xCloseOn, Message := 'ZSC not trusted: still closing at t1 + 59.9 s');
fbTime.Advance(tStep := T#100MS);
fbVlv(itfTime := fbTime, stCmd := stCmd, stRetain := stRetain, stCfg := stCfg);       // t1 + 60 с = tTravel
AssertFalse(Condition := fbVlv.xQClose, Message := 'safe move ends by tTravel');
AssertFalse(Condition := xBoth, Message := 'never both outputs');
fbTime.Advance(tStep := T#1S);
fbVlv(itfTime := fbTime, stCmd := stCmd, stRetain := stRetain, stCfg := stCfg);
AssertFalse(Condition := fbVlv.xQClose, Message := 'not repeated while the interlock stays');
AssertEquals_WORD(Expected := GVL_Const.VLV_FLT_BOTH_LIMITS, Actual := fbVlv.stSts.stCommon.wFault,
                  Message := 'fault still shown');

coUnit.TEST_FINISHED();

(* ---- InterlockWithExtFaultOutputsStayOff.method.decl.st ---- *)
// Авария привода (ExtFault: тепловое реле, обрыв фазы) — привод неисправен: блокировка выходы не включает (VLV-20),
// состояние Fault, бит INTERLOCKED показывает только действующую блокировку.
METHOD PRIVATE InterlockWithExtFaultOutputsStayOff
VAR
    fbTime   : FB_FakeTime;       // подменное время, старт 1 ч
    fbVlv    : FB_Valve;          // арматура под тестом
    stCmd    : ST_ValveCmd;       // команды HMI
    stRetain : ST_DeviceRetain;   // режим, счётчики
    stCfg    : ST_ValveCfg;       // конфигурация (умолчания: Motorized, ZSO и ZSC)
    iStep    : INT;               // шаг цикла

    xAnyOut  : BOOL;              // выход привода хоть раз
END_VAR

(* ---- InterlockWithExtFaultOutputsStayOff.method.impl.st ---- *)
coUnit.TEST('Valve_InterlockWithExtFault_OutputsStayOff');

stRetain.eRemoteMode := E_DeviceMode.Auto;
fbVlv.xAutoOpen := TRUE;
fbVlv.xZso := TRUE;
fbVlv(itfTime := fbTime, stCmd := stCmd, stRetain := stRetain, stCfg := stCfg);       // t0: Open по ZSO
fbVlv.xExtFault := TRUE;
fbTime.Advance(tStep := T#100MS);
fbVlv(itfTime := fbTime, stCmd := stCmd, stRetain := stRetain, stCfg := stCfg);
AssertEquals_WORD(Expected := GVL_Const.VLV_FLT_EXT_FAULT, Actual := fbVlv.stSts.stCommon.wFault,
                  Message := 'precondition: ExtFault');
fbVlv.wInterlock := 16#0001;
FOR iStep := 1 TO 20 DO
    fbTime.Advance(tStep := T#100MS);
    fbVlv(itfTime := fbTime, stCmd := stCmd, stRetain := stRetain, stCfg := stCfg);
    xAnyOut := xAnyOut OR fbVlv.xQOpen OR fbVlv.xQClose;
END_FOR
AssertFalse(Condition := xAnyOut, Message := 'faulty actuator: outputs stay off');
AssertTrue(Condition := fbVlv.stSts.eState = E_ValveState.Fault, Message := 'state Fault');
AssertEquals_WORD(Expected := GVL_Const.VLV_STS_INTERLOCKED,
                  Actual := fbVlv.stSts.stCommon.wStatus AND GVL_Const.VLV_STS_INTERLOCKED,
Message := 'INTERLOCKED bit');

coUnit.TEST_FINISHED();

(* ---- InvalidCfgAtRuntimeKeepsLastValid.method.decl.st ---- *)
// Cfg испорчена в ходе (tTravel = 0): бит wCfgErr и CheckFunction, ход продолжается по последней
// корректной Cfg; время хода контролируется по ней же: FailToOpen ровно на t0 + 10 с.
METHOD PRIVATE InvalidCfgAtRuntimeKeepsLastValid
VAR
    fbTime   : FB_FakeTime;       // подменное время, старт 1 ч
    fbVlv    : FB_Valve;          // арматура под тестом
    stCmd    : ST_ValveCmd;       // команды HMI
    stRetain : ST_DeviceRetain;   // режим Manual по умолчанию, счётчики
    stCfg    : ST_ValveCfg;       // конфигурация (умолчания: Motorized, ZSO и ZSC)
    iStep    : INT;               // шаг цикла
END_VAR

(* ---- InvalidCfgAtRuntimeKeepsLastValid.method.impl.st ---- *)
coUnit.TEST('Valve_InvalidCfgAtRuntime_KeepsLastValid');

stCfg.tTravel := T#10S;
fbVlv.xZsc := TRUE;
fbVlv(itfTime := fbTime, stCmd := stCmd, stRetain := stRetain, stCfg := stCfg);
stCmd.xOpen := TRUE;
// t0
fbVlv(itfTime := fbTime, stCmd := stCmd, stRetain := stRetain, stCfg := stCfg);
fbVlv.xZsc := FALSE;
FOR iStep := 1 TO 20 DO                                                 // t0 + 2,0 с
    fbTime.Advance(tStep := T#100MS);
    fbVlv(itfTime := fbTime, stCmd := stCmd, stRetain := stRetain, stCfg := stCfg);
END_FOR
stCfg.tTravel := T#0S;
fbTime.Advance(tStep := T#100MS);
// t0 + 2,1 с: Cfg испорчена
fbVlv(itfTime := fbTime, stCmd := stCmd, stRetain := stRetain, stCfg := stCfg);
AssertEquals_WORD(Expected := GVL_Const.VLV_CFG_TRAVEL, Actual := fbVlv.stSts.stCommon.wCfgErr, Message := 'wCfgErr');
AssertTrue(Condition := fbVlv.Status = E_Ne107Status.CheckFunction, Message := 'NE 107 CheckFunction');
AssertTrue(Condition := fbVlv.xQOpen, Message := 'keeps running with the last valid cfg');
FOR iStep := 1 TO 78 DO                                                 // t0 + 9,9 с
    fbTime.Advance(tStep := T#100MS);
    fbVlv(itfTime := fbTime, stCmd := stCmd, stRetain := stRetain, stCfg := stCfg);
END_FOR
AssertTrue(Condition := fbVlv.stSts.eState = E_ValveState.Opening, Message := 'Opening at t0 + 9.9 s');
fbTime.Advance(tStep := T#100MS);
// t0 + 10,0 с
fbVlv(itfTime := fbTime, stCmd := stCmd, stRetain := stRetain, stCfg := stCfg);
AssertEquals_WORD(Expected := GVL_Const.VLV_FLT_FAIL_TO_OPEN, Actual := fbVlv.stSts.stCommon.wFault,
                  Message := 'travel supervised with the last valid tTravel');

coUnit.TEST_FINISHED();

(* ---- InvalidCfgStartupOutputsOff.method.decl.st ---- *)
// Корректной Cfg ещё не было (tTravel = T#0S): бит VLV_CFG_TRAVEL, CheckFunction, DEV_STS_CFG_ERROR;
// Auto с запросом «открыть» — выходы сняты 1 с, Available = FALSE; состояние по концевикам; xOpen —
// RejectedCfg без смены режима. Cfg исправлена — арматура идёт к цели.
METHOD PRIVATE InvalidCfgStartupOutputsOff
VAR
    fbTime   : FB_FakeTime;       // подменное время, старт 1 ч
    fbVlv    : FB_Valve;          // арматура под тестом
    stCmd    : ST_ValveCmd;       // команды HMI
    stRetain : ST_DeviceRetain;   // режим Manual по умолчанию, счётчики
    stCfg    : ST_ValveCfg;       // конфигурация (умолчания: Motorized, ZSO и ZSC)
    iStep    : INT;               // шаг цикла
    xEverOn  : BOOL;              // выход включался без корректной Cfg
END_VAR

(* ---- InvalidCfgStartupOutputsOff.method.impl.st ---- *)
coUnit.TEST('Valve_InvalidCfg_StartupOutputsOff');

stCfg.tTravel := T#0S;
stRetain.eRemoteMode := E_DeviceMode.Auto;
fbVlv.xAutoOpen := TRUE;
fbVlv.xZsc := TRUE;
fbVlv(itfTime := fbTime, stCmd := stCmd, stRetain := stRetain, stCfg := stCfg);
AssertEquals_WORD(Expected := GVL_Const.VLV_CFG_TRAVEL, Actual := fbVlv.stSts.stCommon.wCfgErr,
                  Message := 'wCfgErr VLV_CFG_TRAVEL');
AssertTrue(Condition := fbVlv.Status = E_Ne107Status.CheckFunction, Message := 'NE 107 CheckFunction');
AssertEquals_WORD(Expected := GVL_Const.DEV_STS_CFG_ERROR,
                  Actual := fbVlv.stSts.stCommon.wStatus AND GVL_Const.DEV_STS_CFG_ERROR, Message := 'CFG_ERROR bit');
AssertFalse(Condition := fbVlv.Available, Message := 'not available without valid cfg');
FOR iStep := 1 TO 10 DO
    fbTime.Advance(tStep := T#100MS);
    fbVlv(itfTime := fbTime, stCmd := stCmd, stRetain := stRetain, stCfg := stCfg);
    xEverOn := xEverOn OR fbVlv.xQOpen OR fbVlv.xQClose OR fbVlv.xQCoil;
END_FOR
AssertFalse(Condition := xEverOn, Message := 'outputs off without valid cfg');
AssertTrue(Condition := fbVlv.stSts.eState = E_ValveState.Closed, Message := 'state tracks limit switches');
stCmd.xOpen := TRUE;
fbTime.Advance(tStep := T#100MS);
fbVlv(itfTime := fbTime, stCmd := stCmd, stRetain := stRetain, stCfg := stCfg);
AssertTrue(Condition := fbVlv.stSts.stCommon.eCmdResult = E_CmdResult.RejectedCfg, Message := 'RejectedCfg');
AssertTrue(Condition := fbVlv.Mode = E_DeviceMode.Auto, Message := 'rejected command keeps Auto');
stCfg.tTravel := T#60S;
fbTime.Advance(tStep := T#100MS);
fbVlv(itfTime := fbTime, stCmd := stCmd, stRetain := stRetain, stCfg := stCfg);
AssertEquals_WORD(Expected := 0, Actual := fbVlv.stSts.stCommon.wCfgErr, Message := 'cfg valid');
AssertTrue(Condition := fbVlv.xQOpen, Message := 'drives to target once cfg is valid');

coUnit.TEST_FINISHED();

(* ---- LocalOutputsOffTracksLimits.method.decl.st ---- *)
// Local: выходы сняты, команды — RejectedMode; состояние по концевикам при движении руками (цикл
// считается); блокировка — только предупреждение VLV_WRN_INTERLOCK_IN_LOCAL; «оба концевика» не
// контролируется (Unknown, без отказа). Возврат в запомненный Manual без движения.
METHOD PRIVATE LocalOutputsOffTracksLimits
VAR
    fbTime   : FB_FakeTime;       // подменное время, старт 1 ч
    fbVlv    : FB_Valve;          // арматура под тестом
    stCmd    : ST_ValveCmd;       // команды HMI
    stRetain : ST_DeviceRetain;   // режим Manual по умолчанию, счётчики
    stCfg    : ST_ValveCfg;       // конфигурация (умолчания: Motorized, ZSO и ZSC)
    iStep    : INT;               // шаг цикла
END_VAR

(* ---- LocalOutputsOffTracksLimits.method.impl.st ---- *)
coUnit.TEST('Valve_Local_OutputsOffTracksLimits');

fbVlv.xZsc := TRUE;
// Manual, закрыта
fbVlv(itfTime := fbTime, stCmd := stCmd, stRetain := stRetain, stCfg := stCfg);
fbVlv.xLocal := TRUE;
fbVlv(itfTime := fbTime, stCmd := stCmd, stRetain := stRetain, stCfg := stCfg);
AssertTrue(Condition := fbVlv.Mode = E_DeviceMode.Local, Message := 'Local');
stCmd.xOpen := TRUE;
fbVlv(itfTime := fbTime, stCmd := stCmd, stRetain := stRetain, stCfg := stCfg);
AssertTrue(Condition := fbVlv.stSts.stCommon.eCmdResult = E_CmdResult.RejectedMode, Message := 'RejectedMode in Local');
AssertFalse(Condition := fbVlv.xQOpen, Message := 'no output in Local');
fbVlv.xZsc := FALSE;
fbTime.Advance(tStep := T#100MS);
// двигают руками
fbVlv(itfTime := fbTime, stCmd := stCmd, stRetain := stRetain, stCfg := stCfg);
AssertTrue(Condition := fbVlv.stSts.eState = E_ValveState.Intermediate, Message := 'Intermediate between limits');
fbVlv.xZso := TRUE;
fbTime.Advance(tStep := T#100MS);
fbVlv(itfTime := fbTime, stCmd := stCmd, stRetain := stRetain, stCfg := stCfg);
AssertTrue(Condition := fbVlv.stSts.eState = E_ValveState.Open, Message := 'Open on ZSO');
AssertEquals_UDINT(Expected := 1, Actual := stRetain.udiOpCount, Message := 'local cycle counted');
fbVlv.wInterlock := 16#0001;
fbTime.Advance(tStep := T#100MS);
fbVlv(itfTime := fbTime, stCmd := stCmd, stRetain := stRetain, stCfg := stCfg);
AssertEquals_WORD(Expected := GVL_Const.VLV_WRN_INTERLOCK_IN_LOCAL,
                  Actual := fbVlv.stSts.stCommon.wWarning AND GVL_Const.VLV_WRN_INTERLOCK_IN_LOCAL,
                  Message := 'interlock in Local: warning');
AssertEquals_WORD(Expected := 0, Actual := fbVlv.stSts.stCommon.wStatus AND GVL_Const.VLV_STS_INTERLOCKED,
                  Message := 'interlock not acting in Local');
AssertFalse(Condition := fbVlv.xQClose, Message := 'PLC does not move the valve in Local');
fbVlv.xZsc := TRUE;
FOR iStep := 1 TO 10 DO                                                 // оба концевика 1 с
    fbTime.Advance(tStep := T#100MS);
    fbVlv(itfTime := fbTime, stCmd := stCmd, stRetain := stRetain, stCfg := stCfg);
END_FOR
AssertEquals_WORD(Expected := 0, Actual := fbVlv.stSts.stCommon.wFault,
                  Message := 'both limits not supervised in Local');
AssertTrue(Condition := fbVlv.stSts.eState = E_ValveState.Unknown, Message := 'Unknown on both limits');
fbVlv.xZsc := FALSE;
fbVlv.wInterlock := 16#0000;
fbVlv.xLocal := FALSE;
fbTime.Advance(tStep := T#100MS);
fbVlv(itfTime := fbTime, stCmd := stCmd, stRetain := stRetain, stCfg := stCfg);
AssertTrue(Condition := fbVlv.Mode = E_DeviceMode.Manual, Message := 'back to remembered Manual');
AssertTrue(Condition := fbVlv.stSts.eState = E_ValveState.Open, Message := 'Open');
AssertFalse(Condition := fbVlv.xQOpen OR fbVlv.xQClose, Message := 'no movement on return');

coUnit.TEST_FINISHED();

(* ---- MaintCyclesReachedMaintenanceRequired.method.decl.st ---- *)
// ТО по циклам: udiMaintCycles = 2, до ТО остался один цикл. Открытие — счётчик «с ТО» 2: предупреждение
// VLV_WRN_MAINT_CYCLES, NE 107 MaintenanceRequired, бит DEV_STS_WARNING; xResetMaint — снова Good.
METHOD PRIVATE MaintCyclesReachedMaintenanceRequired
VAR
    fbTime   : FB_FakeTime;       // подменное время, старт 1 ч
    fbVlv    : FB_Valve;          // арматура под тестом
    stCmd    : ST_ValveCmd;       // команды HMI
    stRetain : ST_DeviceRetain;   // режим Manual по умолчанию, счётчики
    stCfg    : ST_ValveCfg;       // конфигурация (умолчания: Motorized, ZSO и ZSC)
    iStep    : INT;               // шаг цикла
END_VAR

(* ---- MaintCyclesReachedMaintenanceRequired.method.impl.st ---- *)
coUnit.TEST('Valve_MaintCyclesReached_MaintenanceRequired');

stCfg.udiMaintCycles := 2;
stRetain.udiOpCountMaint := 1;
stRetain.udiOpCount := 41;
fbVlv.xZsc := TRUE;
fbVlv(itfTime := fbTime, stCmd := stCmd, stRetain := stRetain, stCfg := stCfg);
AssertTrue(Condition := fbVlv.Status = E_Ne107Status.Good, Message := 'Good before the interval');
stCmd.xOpen := TRUE;
fbVlv(itfTime := fbTime, stCmd := stCmd, stRetain := stRetain, stCfg := stCfg);
FOR iStep := 1 TO 10 DO
    fbTime.Advance(tStep := T#100MS);
    fbVlv.xZsc := FALSE;
    fbVlv.xZso := iStep >= 10;
    fbVlv(itfTime := fbTime, stCmd := stCmd, stRetain := stRetain, stCfg := stCfg);
END_FOR
AssertEquals_UDINT(Expected := 42, Actual := stRetain.udiOpCount, Message := 'total 42');
AssertEquals_UDINT(Expected := 2, Actual := stRetain.udiOpCountMaint, Message := 'since maintenance 2');
AssertEquals_WORD(Expected := GVL_Const.VLV_WRN_MAINT_CYCLES,
                  Actual := fbVlv.stSts.stCommon.wWarning AND GVL_Const.VLV_WRN_MAINT_CYCLES,
Message := 'MAINT_CYCLES');
AssertTrue(Condition := fbVlv.Status = E_Ne107Status.MaintenanceRequired, Message := 'NE 107 MaintenanceRequired');
AssertEquals_WORD(Expected := GVL_Const.DEV_STS_WARNING,
                  Actual := fbVlv.stSts.stCommon.wStatus AND GVL_Const.DEV_STS_WARNING, Message := 'WARNING bit');
stCmd.xResetMaint := TRUE;
fbTime.Advance(tStep := T#100MS);
fbVlv(itfTime := fbTime, stCmd := stCmd, stRetain := stRetain, stCfg := stCfg);
AssertEquals_UDINT(Expected := 0, Actual := stRetain.udiOpCountMaint, Message := 'reset');
AssertTrue(Condition := fbVlv.Status = E_Ne107Status.Good, Message := 'Good after maintenance reset');
AssertEquals_UDINT(Expected := 42, Actual := stRetain.udiOpCount, Message := 'total kept');

coUnit.TEST_FINISHED();

(* ---- ManualCmdInAutoSwitchesToManual.method.decl.st ---- *)
// Auto, запрос «закрыть», закрыта. xOpen оператора: Manual (запоминается в stRetain), Opening, Accepted;
// запрос автоматики больше не действует. xStop в Auto: Manual и стоп.
METHOD PRIVATE ManualCmdInAutoSwitchesToManual
VAR
    fbTime   : FB_FakeTime;       // подменное время, старт 1 ч
    fbVlv    : FB_Valve;          // арматура под тестом
    stCmd    : ST_ValveCmd;       // команды HMI
    stRetain : ST_DeviceRetain;   // режим Manual по умолчанию, счётчики
    stCfg    : ST_ValveCfg;       // конфигурация (умолчания: Motorized, ZSO и ZSC)
END_VAR

(* ---- NeverBothOutputs.method.decl.st ---- *)
// Инвариант: xQOpen AND xQClose никогда не TRUE. 600 циклов по 0,1 с с моделью хода (30 шагов от ZSC до
// ZSO): команды открыть, закрыть, стоп с разными периодами, переходы в Auto с переменным запросом,
// блокировки и пропадающее разрешение на открытие. Проверяется и то, что сценарий открывал, закрывал и
// реверсировал (тест не пустой).
METHOD PRIVATE NeverBothOutputs
VAR
    fbTime    : FB_FakeTime;       // подменное время, старт 1 ч
    fbVlv     : FB_Valve;          // арматура под тестом
    stCmd     : ST_ValveCmd;       // команды HMI
    stRetain  : ST_DeviceRetain;   // режим Manual по умолчанию, счётчики
    stCfg     : ST_ValveCfg;       // конфигурация (умолчания: Motorized, ZSO и ZSC)
    iStep     : INT;               // шаг цикла
    iPos      : INT;               // положение модели, шаги 0…30
    xEverBoth : BOOL;              // оба выхода хоть раз
    xSawOpen  : BOOL;              // открывала
    xSawClose : BOOL;              // закрывала
    xSawRev   : BOOL;              // реверсировала
END_VAR

(* ---- NeverBothOutputs.method.impl.st ---- *)
coUnit.TEST('Valve_NeverBothOutputs');

stCfg.tTravel := T#5S;
stCfg.tReverse := T#300MS;
fbVlv.xZsc := TRUE;
fbVlv(itfTime := fbTime, stCmd := stCmd, stRetain := stRetain, stCfg := stCfg);
FOR iStep := 1 TO 600 DO
    fbTime.Advance(tStep := T#100MS);
    IF fbVlv.xQOpen THEN
        iPos := iPos + 1;
    END_IF
    IF fbVlv.xQClose THEN
        iPos := iPos - 1;
    END_IF
    iPos := LIMIT(0, iPos, 30);
    fbVlv.xZso := iPos >= 30;
    fbVlv.xZsc := iPos <= 0;
    stCmd.xOpen := iStep MOD 11 = 0;
    stCmd.xClose := iStep MOD 7 = 0;
    stCmd.xStop := iStep MOD 23 = 0;
    stCmd.stCommon.xSetAuto := iStep MOD 97 = 0;
    fbVlv.xAutoOpen := (iStep / 13) MOD 2 = 0;
    fbVlv.wInterlock := SEL((iStep / 40) MOD 4 = 3, 16#0000, 16#0001);
    fbVlv.wPermitOpen := SEL((iStep / 60) MOD 3 = 1, 16#FFFF, 16#0000);
    fbVlv(itfTime := fbTime, stCmd := stCmd, stRetain := stRetain, stCfg := stCfg);
    xEverBoth := xEverBoth OR (fbVlv.xQOpen AND fbVlv.xQClose);
    xSawOpen := xSawOpen OR fbVlv.xQOpen;
    xSawClose := xSawClose OR fbVlv.xQClose;
    xSawRev := xSawRev OR fbVlv.stSts.eState = E_ValveState.Reversing;
END_FOR
AssertFalse(Condition := xEverBoth, Message := 'never both contactors');
AssertTrue(Condition := xSawOpen, Message := 'scenario opened');
AssertTrue(Condition := xSawClose, Message := 'scenario closed');
AssertTrue(Condition := xSawRev, Message := 'scenario reversed');

coUnit.TEST_FINISHED();

(* ---- NoLimitSwitchesPositionByTravelTime.method.decl.st ---- *)
// Концевиков нет: старт — Unknown (VLV_WRN_POSITION_UNKNOWN). xOpen: выход держится tTravel = 10 с (на
// 9,9 с ещё Opening), ровно на 10,0 с — Open по времени без отказа, VLV_WRN_POSITION_BY_TIME; входы
// неподключённых концевиков не учитываются.
METHOD PRIVATE NoLimitSwitchesPositionByTravelTime
VAR
    fbTime   : FB_FakeTime;       // подменное время, старт 1 ч
    fbVlv    : FB_Valve;          // арматура под тестом
    stCmd    : ST_ValveCmd;       // команды HMI
    stRetain : ST_DeviceRetain;   // режим Manual по умолчанию, счётчики
    stCfg    : ST_ValveCfg;       // конфигурация (умолчания: Motorized, ZSO и ZSC)
    iStep    : INT;               // шаг цикла
END_VAR

(* ---- NoLimitSwitchesPositionByTravelTime.method.impl.st ---- *)
coUnit.TEST('Valve_NoLimitSwitches_PositionByTravelTime');

stCfg.xZsoUsed := FALSE;
stCfg.xZscUsed := FALSE;
stCfg.tTravel := T#10S;
fbVlv(itfTime := fbTime, stCmd := stCmd, stRetain := stRetain, stCfg := stCfg);
AssertTrue(Condition := fbVlv.stSts.eState = E_ValveState.Unknown, Message := 'Unknown without limit switches');
AssertEquals_WORD(Expected := GVL_Const.VLV_WRN_POSITION_UNKNOWN,
                  Actual := fbVlv.stSts.stCommon.wWarning AND GVL_Const.VLV_WRN_POSITION_UNKNOWN,
                  Message := 'POSITION_UNKNOWN warning');
stCmd.xOpen := TRUE;
// t0
fbVlv(itfTime := fbTime, stCmd := stCmd, stRetain := stRetain, stCfg := stCfg);
FOR iStep := 1 TO 99 DO                                                 // t0 + 9,9 с
    fbTime.Advance(tStep := T#100MS);
    fbVlv(itfTime := fbTime, stCmd := stCmd, stRetain := stRetain, stCfg := stCfg);
END_FOR
AssertTrue(Condition := fbVlv.stSts.eState = E_ValveState.Opening, Message := 'Opening at t0 + 9.9 s');
AssertTrue(Condition := fbVlv.xQOpen, Message := 'output held until tTravel');
fbTime.Advance(tStep := T#100MS);
// t0 + 10,0 с
fbVlv(itfTime := fbTime, stCmd := stCmd, stRetain := stRetain, stCfg := stCfg);
AssertTrue(Condition := fbVlv.stSts.eState = E_ValveState.Open, Message := 'Open by travel time');
AssertFalse(Condition := fbVlv.xQOpen, Message := 'output off');
AssertTrue(Condition := fbVlv.xOpened, Message := 'xOpened');
AssertEquals_WORD(Expected := 0, Actual := fbVlv.stSts.stCommon.wFault, Message := 'no fault without limit switch');
AssertEquals_WORD(Expected := GVL_Const.VLV_WRN_POSITION_BY_TIME,
                  Actual := fbVlv.stSts.stCommon.wWarning AND GVL_Const.VLV_WRN_POSITION_BY_TIME,
                  Message := 'POSITION_BY_TIME warning');
fbVlv.xZsc := TRUE;
fbTime.Advance(tStep := T#100MS);
fbVlv(itfTime := fbTime, stCmd := stCmd, stRetain := stRetain, stCfg := stCfg);
AssertTrue(Condition := fbVlv.stSts.eState = E_ValveState.Open, Message := 'unused ZSC ignored');

coUnit.TEST_FINISHED();

(* ---- OosEntryClearsLatchedFaults.method.decl.st ---- *)
// Зафиксированные TorqueTrip (муфта в ходе после страгивания, отпустила) и внешняя авария (причина ушла)
// снимаются входом в OutOfService; в OOS внешняя авария не контролируется, тревоги — OutOfService; после выхода
// в Manual отказа нет.
METHOD PRIVATE OosEntryClearsLatchedFaults
VAR
    fbTime   : FB_FakeTime;       // подменное время, старт 1 ч
    fbVlv    : FB_Valve;          // арматура под тестом
    stCmd    : ST_ValveCmd;       // команды HMI
    stRetain : ST_DeviceRetain;   // режим Manual по умолчанию, счётчики
    stCfg    : ST_ValveCfg;       // конфигурация (умолчания: Motorized, ZSO и ZSC)
    itfAlm   : I_Alarm;           // слот тревоги через интерфейс
END_VAR

(* ---- OosRequestWhileMovingRejected.method.decl.st ---- *)
// Вывод из работы в ходе — RejectedState, ход продолжается. Остановленную арматуру вывести можно:
// OutOfService, выходы сняты, CheckFunction, команды — RejectedMode.
METHOD PRIVATE OosRequestWhileMovingRejected
VAR
    fbTime   : FB_FakeTime;       // подменное время, старт 1 ч
    fbVlv    : FB_Valve;          // арматура под тестом
    stCmd    : ST_ValveCmd;       // команды HMI
    stRetain : ST_DeviceRetain;   // режим Manual по умолчанию, счётчики
    stCfg    : ST_ValveCfg;       // конфигурация (умолчания: Motorized, ZSO и ZSC)
END_VAR

(* ---- OpenLimitReachedGoesOpen.method.decl.st ---- *)
// Manual, задвижка закрыта (ZSC). xOpen: Opening, включён только xQOpen, остаток хода 10 с; через 2 с
// остаток 8 с; ZSO на t0 + 5,0 с — Open, выход снят, xOpened, один цикл в stRetain.
METHOD PRIVATE OpenLimitReachedGoesOpen
VAR
    fbTime   : FB_FakeTime;       // подменное время, старт 1 ч
    fbVlv    : FB_Valve;          // арматура под тестом
    stCmd    : ST_ValveCmd;       // команды HMI
    stRetain : ST_DeviceRetain;   // режим Manual по умолчанию, счётчики
    stCfg    : ST_ValveCfg;       // конфигурация (умолчания: Motorized, ZSO и ZSC)
    iStep    : INT;               // шаг цикла
END_VAR

(* ---- OpenLimitReachedGoesOpen.method.impl.st ---- *)
coUnit.TEST('Valve_Open_LimitReached_GoesOpen');

stCfg.tTravel := T#10S;
fbVlv.xZsc := TRUE;
// t0: закрыта
fbVlv(itfTime := fbTime, stCmd := stCmd, stRetain := stRetain, stCfg := stCfg);
AssertTrue(Condition := fbVlv.stSts.eState = E_ValveState.Closed, Message := 'starts Closed on ZSC');
AssertTrue(Condition := fbVlv.xClosed, Message := 'xClosed on ZSC');
stCmd.xOpen := TRUE;
// t0: команда «открыть»
fbVlv(itfTime := fbTime, stCmd := stCmd, stRetain := stRetain, stCfg := stCfg);
AssertTrue(Condition := fbVlv.stSts.eState = E_ValveState.Opening, Message := 'Opening after xOpen');
AssertTrue(Condition := fbVlv.xQOpen, Message := 'open contactor on');
AssertFalse(Condition := fbVlv.xQClose, Message := 'close contactor off');
AssertFalse(Condition := stCmd.xOpen, Message := 'xOpen cleared');
AssertTrue(Condition := fbVlv.stSts.stCommon.eCmdResult = E_CmdResult.Accepted, Message := 'open accepted');
// источник: tools/reference/valve_reference.py, сценарий valve_travel_remain (elapsed 0 s)
AssertEquals_UINT(Expected := 10, Actual := fbVlv.stSts.uiTravelRemain_s, Message := 'travel remain 10 s at start');
FOR iStep := 1 TO 20 DO                                                 // t0 + 0,1 … 2,0 с; ZSC пропал на 0,5 с
    fbTime.Advance(tStep := T#100MS);
    fbVlv.xZsc := iStep < 5;
    fbVlv(itfTime := fbTime, stCmd := stCmd, stRetain := stRetain, stCfg := stCfg);
END_FOR
// источник: tools/reference/valve_reference.py, сценарий valve_travel_remain (elapsed 2.0 s)
AssertEquals_UINT(Expected := 8, Actual := fbVlv.stSts.uiTravelRemain_s, Message := 'travel remain 8 s at t0 + 2 s');
AssertEquals_WORD(Expected := GVL_Const.VLV_STS_OPENING,
                  Actual := fbVlv.stSts.stCommon.wStatus AND GVL_Const.VLV_STS_OPENING, Message := 'OPENING bit');
FOR iStep := 21 TO 49 DO                                                // до t0 + 4,9 с
    fbTime.Advance(tStep := T#100MS);
    fbVlv(itfTime := fbTime, stCmd := stCmd, stRetain := stRetain, stCfg := stCfg);
END_FOR
AssertTrue(Condition := fbVlv.xQOpen, Message := 'still opening at t0 + 4.9 s');
fbTime.Advance(tStep := T#100MS);
fbVlv.xZso := TRUE;
// t0 + 5,0 с: ZSO
fbVlv(itfTime := fbTime, stCmd := stCmd, stRetain := stRetain, stCfg := stCfg);
AssertTrue(Condition := fbVlv.stSts.eState = E_ValveState.Open, Message := 'Open on ZSO');
AssertFalse(Condition := fbVlv.xQOpen, Message := 'contactor off at ZSO');
AssertTrue(Condition := fbVlv.xOpened, Message := 'xOpened');
AssertEquals_WORD(Expected := GVL_Const.VLV_STS_OPENED,
                  Actual := fbVlv.stSts.stCommon.wStatus
                            AND (GVL_Const.VLV_STS_OPENED OR GVL_Const.VLV_STS_CLOSED OR GVL_Const.VLV_STS_OPENING),
                  Message := 'only OPENED of the position bits');
AssertEquals_UDINT(Expected := 1, Actual := stRetain.udiOpCount, Message := 'one open cycle counted');
AssertEquals_UINT(Expected := 0, Actual := fbVlv.stSts.uiTravelRemain_s, Message := 'no travel remain at rest');
AssertEquals_WORD(Expected := 0, Actual := fbVlv.stSts.stCommon.wFault, Message := 'no fault');

coUnit.TEST_FINISHED();

(* ---- OpenTimeoutSetsFailToOpen.method.decl.st ---- *)
// tTravel = 10 с, ZSO не приходит: на t0 + 9,9 с ещё Opening без отказа, ровно на t0 + 10,0 с —
// FailToOpen (wFault бит 0, Failure, тревога слота 0), выход снят. Отказ фиксируется: пришедший позже
// ZSO его не снимает (положение видно в xOpened), снимает Reset — далее состояние по концевикам.
METHOD PRIVATE OpenTimeoutSetsFailToOpen
VAR
    fbTime   : FB_FakeTime;       // подменное время, старт 1 ч
    fbVlv    : FB_Valve;          // арматура под тестом
    stCmd    : ST_ValveCmd;       // команды HMI
    stRetain : ST_DeviceRetain;   // режим Manual по умолчанию, счётчики
    stCfg    : ST_ValveCfg;       // конфигурация (умолчания: Motorized, ZSO и ZSC)
    iStep    : INT;               // шаг цикла
    itfAlm   : I_Alarm;           // слот тревоги через интерфейс
END_VAR

(* ---- OpenTimeoutSetsFailToOpen.method.impl.st ---- *)
coUnit.TEST('Valve_Open_Timeout_SetsFailToOpen');

stCfg.tTravel := T#10S;
fbVlv.xZsc := TRUE;
// t0: закрыта
fbVlv(itfTime := fbTime, stCmd := stCmd, stRetain := stRetain, stCfg := stCfg);
stCmd.xOpen := TRUE;
// t0: Opening
fbVlv(itfTime := fbTime, stCmd := stCmd, stRetain := stRetain, stCfg := stCfg);
fbVlv.xZsc := FALSE;
FOR iStep := 1 TO 99 DO                                                 // до t0 + 9,9 с ZSO нет
    fbTime.Advance(tStep := T#100MS);
    fbVlv(itfTime := fbTime, stCmd := stCmd, stRetain := stRetain, stCfg := stCfg);
END_FOR
AssertTrue(Condition := fbVlv.stSts.eState = E_ValveState.Opening, Message := 'still opening at t0 + 9.9 s');
AssertEquals_WORD(Expected := 0, Actual := fbVlv.stSts.stCommon.wFault, Message := 'no fault before tTravel');
fbTime.Advance(tStep := T#100MS);
// t0 + 10,0 с
fbVlv(itfTime := fbTime, stCmd := stCmd, stRetain := stRetain, stCfg := stCfg);
AssertTrue(Condition := fbVlv.stSts.eState = E_ValveState.Fault, Message := 'Fault at tTravel');
AssertFalse(Condition := fbVlv.xQOpen, Message := 'output off on timeout');
AssertEquals_WORD(Expected := GVL_Const.VLV_FLT_FAIL_TO_OPEN, Actual := fbVlv.stSts.stCommon.wFault,
                  Message := 'wFault FailToOpen');
AssertTrue(Condition := fbVlv.Status = E_Ne107Status.Failure, Message := 'NE 107 Failure');
itfAlm := fbVlv.GetAlarm(uiIndex := E_ValveAlarm.FailToOpen);
AssertTrue(Condition := itfAlm.State = E_AlarmState.ActiveUnack, Message := 'FailToOpen alarm ActiveUnack');
fbTime.Advance(tStep := T#100MS);
fbVlv.xZso := TRUE;
// ZSO пришёл позже
fbVlv(itfTime := fbTime, stCmd := stCmd, stRetain := stRetain, stCfg := stCfg);
AssertEquals_WORD(Expected := GVL_Const.VLV_FLT_FAIL_TO_OPEN, Actual := fbVlv.stSts.stCommon.wFault,
                  Message := 'fault latched');
AssertTrue(Condition := fbVlv.xOpened, Message := 'position still visible in Fault');
stCmd.stCommon.xReset := TRUE;
fbVlv(itfTime := fbTime, stCmd := stCmd, stRetain := stRetain, stCfg := stCfg);
AssertTrue(Condition := fbVlv.stSts.stCommon.eCmdResult = E_CmdResult.Accepted, Message := 'Reset accepted');
AssertEquals_WORD(Expected := 0, Actual := fbVlv.stSts.stCommon.wFault, Message := 'cleared by Reset');
AssertTrue(Condition := fbVlv.stSts.eState = E_ValveState.Open, Message := 'state from limit switches after Reset');
AssertFalse(Condition := fbVlv.xQOpen, Message := 'no output after Reset');

coUnit.TEST_FINISHED();

(* ---- OpenTorqueUnseatingNoZscTripsAfterBypass.method.decl.st ---- *)
// Закрытие по моменту без ZSC (xZscUsed = FALSE): задвижка закрыта по муфте. «Открыть»: муфта открытия держится —
// при страгивании с закрытого положения она не контролируется VLV_UNSEAT_BYPASS = 2 с от начала хода (VLV-21);
// держится дольше — клин не вышел из седла: TorqueTrip ровно через 2 с, выход снят.
METHOD PRIVATE OpenTorqueUnseatingNoZscTripsAfterBypass
VAR
    fbTime   : FB_FakeTime;       // подменное время, старт 1 ч
    fbVlv    : FB_Valve;          // арматура под тестом
    stCmd    : ST_ValveCmd;       // команды HMI
    stRetain : ST_DeviceRetain;   // режим, счётчики
    stCfg    : ST_ValveCfg;       // конфигурация (умолчания: Motorized, ZSO и ZSC)
    iStep    : INT;               // шаг цикла
END_VAR

(* ---- OpenTorqueUnseatingNoZscTripsAfterBypass.method.impl.st ---- *)
coUnit.TEST('Valve_OpenTorqueUnseatingNoZsc_TripsAfterBypass');

stCfg.xZscUsed := FALSE;
stCfg.xTorqueUsed := TRUE;
stCfg.xCloseOnTorque := TRUE;
fbVlv(itfTime := fbTime, stCmd := stCmd, stRetain := stRetain, stCfg := stCfg);       // t0
stCmd.xClose := TRUE;
fbTime.Advance(tStep := T#100MS);
fbVlv(itfTime := fbTime, stCmd := stCmd, stRetain := stRetain, stCfg := stCfg);       // Closing
fbVlv.xTorqueClose := TRUE;
fbTime.Advance(tStep := T#100MS);
fbVlv(itfTime := fbTime, stCmd := stCmd, stRetain := stRetain, stCfg := stCfg);       // посадка по муфте
AssertTrue(Condition := fbVlv.stSts.eState = E_ValveState.Closed, Message := 'precondition: closed on torque');
fbVlv.xTorqueClose := FALSE;
fbTime.Advance(tStep := T#2S);
fbVlv(itfTime := fbTime, stCmd := stCmd, stRetain := stRetain, stCfg := stCfg);       // выбег прошёл (tReverse)
stCmd.xOpen := TRUE;
fbVlv.xTorqueOpen := TRUE;
fbTime.Advance(tStep := T#100MS);
fbVlv(itfTime := fbTime, stCmd := stCmd, stRetain := stRetain, stCfg := stCfg);   // t1: Opening с седла, муфта сразу
AssertTrue(Condition := fbVlv.xQOpen, Message := 'precondition: opening from the seat');
FOR iStep := 1 TO 19 DO
    fbTime.Advance(tStep := T#100MS);
    fbVlv(itfTime := fbTime, stCmd := stCmd, stRetain := stRetain, stCfg := stCfg);
END_FOR
AssertTrue(Condition := fbVlv.xQOpen, Message := 'torque ignored within the unseating bypass (1.9 s)');
AssertEquals_WORD(Expected := 0, Actual := fbVlv.stSts.stCommon.wFault, Message := 'no fault within the bypass');
fbTime.Advance(tStep := T#100MS);
fbVlv(itfTime := fbTime, stCmd := stCmd, stRetain := stRetain, stCfg := stCfg);       // t1 + 2,0 с
AssertEquals_WORD(Expected := GVL_Const.VLV_FLT_TORQUE_TRIP, Actual := fbVlv.stSts.stCommon.wFault,
                  Message := 'TorqueTrip exactly at the end of the bypass');
AssertFalse(Condition := fbVlv.xQOpen, Message := 'output off');

coUnit.TEST_FINISHED();

(* ---- OpenTorqueWhileUnseatingIgnored.method.decl.st ---- *)
// Клиновая задвижка, закрытие по моменту (xTorqueUsed, xCloseOnTorque), закрыта при ZSC. «Открыть»: при страгивании
// клина муфта открытия срабатывает, пока ZSC ещё замкнут, — это не заклинивание (VLV-21): ход продолжается, отказа
// нет. ZSC разомкнулся; ещё tLimitFilter (0,5 с) муфта не контролируется, затем муфта в ходе — TorqueTrip.
METHOD PRIVATE OpenTorqueWhileUnseatingIgnored
VAR
    fbTime   : FB_FakeTime;       // подменное время, старт 1 ч
    fbVlv    : FB_Valve;          // арматура под тестом
    stCmd    : ST_ValveCmd;       // команды HMI
    stRetain : ST_DeviceRetain;   // режим, счётчики
    stCfg    : ST_ValveCfg;       // конфигурация (умолчания: Motorized, ZSO и ZSC)
    iStep    : INT;               // шаг цикла
END_VAR

(* ---- OpenTorqueWhileUnseatingIgnored.method.impl.st ---- *)
coUnit.TEST('Valve_OpenTorqueWhileUnseating_Ignored');

stCfg.xTorqueUsed := TRUE;
stCfg.xCloseOnTorque := TRUE;
fbVlv.xZsc := TRUE;
fbVlv(itfTime := fbTime, stCmd := stCmd, stRetain := stRetain, stCfg := stCfg);       // t0: Closed по ZSC (старт ПЛК)
AssertTrue(Condition := fbVlv.stSts.eState = E_ValveState.Closed, Message := 'precondition: Closed');
stCmd.xOpen := TRUE;
fbTime.Advance(tStep := T#100MS);
fbVlv(itfTime := fbTime, stCmd := stCmd, stRetain := stRetain, stCfg := stCfg);       // t1: Opening
AssertTrue(Condition := fbVlv.xQOpen, Message := 'precondition: opening');
fbVlv.xTorqueOpen := TRUE;                                                             // страгивание клина
FOR iStep := 1 TO 3 DO
    fbTime.Advance(tStep := T#100MS);
    fbVlv(itfTime := fbTime, stCmd := stCmd, stRetain := stRetain, stCfg := stCfg);
END_FOR
AssertTrue(Condition := fbVlv.xQOpen, Message := 'unseating torque ignored while ZSC is made');
AssertEquals_WORD(Expected := 0, Actual := fbVlv.stSts.stCommon.wFault, Message := 'no TorqueTrip at unseating');
fbVlv.xZsc := FALSE;                                                                   // t1 + 0,4 с: клин вышел
FOR iStep := 1 TO 5 DO                                                               // t1 + 0,4 … t1 + 0,8 с
    fbTime.Advance(tStep := T#100MS);
    fbVlv(itfTime := fbTime, stCmd := stCmd, stRetain := stRetain, stCfg := stCfg);
END_FOR
AssertTrue(Condition := fbVlv.xQOpen, Message := 'bypass held for tLimitFilter after ZSC released');
fbTime.Advance(tStep := T#100MS);
fbVlv(itfTime := fbTime, stCmd := stCmd, stRetain := stRetain, stCfg := stCfg);       // t1 + 0,9 с: ZSC разомкнут 0,5 с
AssertEquals_WORD(Expected := GVL_Const.VLV_FLT_TORQUE_TRIP, Actual := fbVlv.stSts.stCommon.wFault,
                  Message := 'torque after unseating trips');
AssertFalse(Condition := fbVlv.xQOpen, Message := 'output off');

coUnit.TEST_FINISHED();

(* ---- PermitCloseMissingAutoWaitsReportsCloseBits.method.decl.st ---- *)
// Auto, задвижка открыта. Нет разрешения на закрытие (бит 1), а на открытие не хватает другого бита
// (бит 0). Автоматика просит «закрыть»: выход «закрывать» не включается, бит PERMIT_MISSING, в
// wPermitMissing — недостающие биты направления к цели (16#0002), а не открытия. Разрешение появилось —
// задвижка закрывается, wPermitMissing = 0.
METHOD PRIVATE PermitCloseMissingAutoWaitsReportsCloseBits
VAR
    fbTime   : FB_FakeTime;       // подменное время, старт 1 ч
    fbVlv    : FB_Valve;          // арматура под тестом
    stCmd    : ST_ValveCmd;       // команды HMI
    stRetain : ST_DeviceRetain;   // режим: Auto
    stCfg    : ST_ValveCfg;       // конфигурация (умолчания: Motorized, ZSO и ZSC)
END_VAR

(* ---- PermitLostWhileMovingContinuesMotion.method.decl.st ---- *)
// Разрешение на открытие пропало в ходе: работающий ход не останавливается (бит PERMIT_MISSING и
// wPermitMissing показывают недостачу), арматура доходит до ZSO.
METHOD PRIVATE PermitLostWhileMovingContinuesMotion
VAR
    fbTime   : FB_FakeTime;       // подменное время, старт 1 ч
    fbVlv    : FB_Valve;          // арматура под тестом
    stCmd    : ST_ValveCmd;       // команды HMI
    stRetain : ST_DeviceRetain;   // режим Manual по умолчанию, счётчики
    stCfg    : ST_ValveCfg;       // конфигурация (умолчания: Motorized, ZSO и ZSC)
    iStep    : INT;               // шаг цикла
END_VAR

(* ---- PermitLostWhileMovingContinuesMotion.method.impl.st ---- *)
coUnit.TEST('Valve_PermitLostWhileMoving_ContinuesMotion');

fbVlv.xZsc := TRUE;
fbVlv(itfTime := fbTime, stCmd := stCmd, stRetain := stRetain, stCfg := stCfg);
stCmd.xOpen := TRUE;
fbVlv(itfTime := fbTime, stCmd := stCmd, stRetain := stRetain, stCfg := stCfg);
fbVlv.xZsc := FALSE;
FOR iStep := 1 TO 10 DO
    fbTime.Advance(tStep := T#100MS);
    fbVlv(itfTime := fbTime, stCmd := stCmd, stRetain := stRetain, stCfg := stCfg);
END_FOR
fbVlv.wPermitOpen := 16#0000;
fbTime.Advance(tStep := T#100MS);
fbVlv(itfTime := fbTime, stCmd := stCmd, stRetain := stRetain, stCfg := stCfg);
AssertTrue(Condition := fbVlv.xQOpen, Message := 'running stroke not stopped by a lost permit');
AssertEquals_WORD(Expected := GVL_Const.VLV_STS_PERMIT_MISSING,
                  Actual := fbVlv.stSts.stCommon.wStatus AND GVL_Const.VLV_STS_PERMIT_MISSING,
                  Message := 'PERMIT_MISSING bit');
AssertEquals_WORD(Expected := 16#FFFF, Actual := fbVlv.stSts.wPermitMissing, Message := 'all open permits missing');
FOR iStep := 1 TO 10 DO
    fbTime.Advance(tStep := T#100MS);
    fbVlv.xZso := iStep >= 10;
    fbVlv(itfTime := fbTime, stCmd := stCmd, stRetain := stRetain, stCfg := stCfg);
END_FOR
AssertTrue(Condition := fbVlv.stSts.eState = E_ValveState.Open, Message := 'reaches Open');

coUnit.TEST_FINISHED();

(* ---- PermitOpenMissingOpenRejected.method.decl.st ---- *)
// Нет разрешения на открытие (бит 0): xOpen — RejectedPermit, движения нет; бит снят из маски —
// команда принята. В Auto запрос «открыть» ждёт разрешения (бит PERMIT_MISSING, wPermitMissing) и
// выполняется, когда оно появится.
METHOD PRIVATE PermitOpenMissingOpenRejected
VAR
    fbTime   : FB_FakeTime;       // подменное время, старт 1 ч
    fbVlv    : FB_Valve;          // арматура под тестом
    stCmd    : ST_ValveCmd;       // команды HMI
    stRetain : ST_DeviceRetain;   // режим Manual по умолчанию, счётчики
    stCfg    : ST_ValveCfg;       // конфигурация (умолчания: Motorized, ZSO и ZSC)
END_VAR

(* ---- PlcRestartStateFromLimits.method.decl.st ---- *)
// Старт ПЛК (первый вызов, Manual): ZSO — Open, оба концевика — сразу Fault (BothLimits), ни одного —
// Intermediate, без концевиков — Unknown; выходы сняты.
METHOD PRIVATE PlcRestartStateFromLimits
VAR
    fbTime    : FB_FakeTime;       // подменное время
    fbOpen    : FB_Valve;          // старт на ZSO
    fbBoth    : FB_Valve;          // старт на обоих концевиках
    fbMid     : FB_Valve;          // старт без сигналов концевиков
    fbNone    : FB_Valve;          // старт без подключённых концевиков
    stCmd     : ST_ValveCmd;       // команды (общие: пустые)
    stRetain  : ST_DeviceRetain;   // Manual
    stCfg     : ST_ValveCfg;       // умолчания
    stCfgNone : ST_ValveCfg;       // концевики не подключены
END_VAR

(* ---- PositionByTimeLostInLocalAutoDrivesAgain.method.decl.st ---- *)
// Концевиков нет, Auto: открыта по времени хода (tTravel = 10 с, на t0 + 10,0 с — Open). Local: с места
// арматуру могут закрыть, положение «по времени» больше не известно — Unknown, xOpened нет,
// VLV_WRN_POSITION_UNKNOWN. Возврат в дистанционный режим (Auto, xAutoOpen): привод снова ведёт к цели —
// Opening, выход «открывать» на tTravel, ровно через 10,0 с — снова Open по времени. С устаревшим «Open»
// автоматика считала бы открытой задвижку, которую закрыли с места.
METHOD PRIVATE PositionByTimeLostInLocalAutoDrivesAgain
VAR
    fbTime   : FB_FakeTime;       // подменное время, старт 1 ч
    fbVlv    : FB_Valve;          // арматура под тестом
    stCmd    : ST_ValveCmd;       // команды HMI
    stRetain : ST_DeviceRetain;   // режим: Auto
    stCfg    : ST_ValveCfg;       // конфигурация: без концевиков
    iStep    : INT;               // шаг цикла
END_VAR

(* ---- PositionByTimeLostInLocalAutoDrivesAgain.method.impl.st ---- *)
coUnit.TEST('Valve_PositionByTime_LostInLocal_AutoDrivesAgain');

stCfg.xZsoUsed := FALSE;
stCfg.xZscUsed := FALSE;
stCfg.tTravel := T#10S;
stRetain.eRemoteMode := E_DeviceMode.Auto;
fbVlv.xAutoOpen := TRUE;
// t0: Auto ведёт к цели
fbVlv(itfTime := fbTime, stCmd := stCmd, stRetain := stRetain, stCfg := stCfg);
AssertTrue(Condition := fbVlv.xQOpen, Message := 'Auto opens');
FOR iStep := 1 TO 100 DO                                                // t0 + 10,0 с
    fbTime.Advance(tStep := T#100MS);
    fbVlv(itfTime := fbTime, stCmd := stCmd, stRetain := stRetain, stCfg := stCfg);
END_FOR
AssertTrue(Condition := fbVlv.stSts.eState = E_ValveState.Open, Message := 'Open by travel time');
AssertTrue(Condition := fbVlv.xOpened, Message := 'xOpened by time');
fbVlv.xLocal := TRUE;
fbTime.Advance(tStep := T#100MS);
fbVlv(itfTime := fbTime, stCmd := stCmd, stRetain := stRetain, stCfg := stCfg);
AssertTrue(Condition := fbVlv.Mode = E_DeviceMode.Local, Message := 'Local');
AssertTrue(Condition := fbVlv.stSts.eState = E_ValveState.Unknown, Message := 'position by time lost in Local');
AssertFalse(Condition := fbVlv.xOpened, Message := 'not reported open in Local');
AssertEquals_WORD(Expected := GVL_Const.VLV_WRN_POSITION_UNKNOWN,
                  Actual := fbVlv.stSts.stCommon.wWarning AND GVL_Const.VLV_WRN_POSITION_UNKNOWN,
                  Message := 'POSITION_UNKNOWN warning');
FOR iStep := 1 TO 50 DO                                                 // 5 с в Local
    fbTime.Advance(tStep := T#100MS);
    fbVlv(itfTime := fbTime, stCmd := stCmd, stRetain := stRetain, stCfg := stCfg);
END_FOR
fbVlv.xLocal := FALSE;
fbTime.Advance(tStep := T#100MS);
// t1: снова Auto
fbVlv(itfTime := fbTime, stCmd := stCmd, stRetain := stRetain, stCfg := stCfg);
AssertTrue(Condition := fbVlv.Mode = E_DeviceMode.Auto, Message := 'back to Auto');
AssertTrue(Condition := fbVlv.stSts.eState = E_ValveState.Opening, Message := 'Auto drives to target again');
AssertTrue(Condition := fbVlv.xQOpen, Message := 'open contactor on');
FOR iStep := 1 TO 99 DO                                                 // t1 + 9,9 с
    fbTime.Advance(tStep := T#100MS);
    fbVlv(itfTime := fbTime, stCmd := stCmd, stRetain := stRetain, stCfg := stCfg);
END_FOR
AssertTrue(Condition := fbVlv.stSts.eState = E_ValveState.Opening, Message := 'Opening at t1 + 9.9 s');
fbTime.Advance(tStep := T#100MS);
// t1 + 10,0 с
fbVlv(itfTime := fbTime, stCmd := stCmd, stRetain := stRetain, stCfg := stCfg);
AssertTrue(Condition := fbVlv.stSts.eState = E_ValveState.Open, Message := 'Open by travel time again');
AssertEquals_WORD(Expected := 0, Actual := fbVlv.stSts.stCommon.wFault, Message := 'no fault');

coUnit.TEST_FINISHED();

(* ---- PositionLostLatchesFault.method.decl.st ---- *)
// Manual, открыта. Провал ZSO на 0,4 с фильтруется (tLimitFilter = 0,5 с). Пропал на 0,5 с без команды —
// PositionLost (wFault бит 3), фиксируется: вернувшийся ZSO отказ не снимает, снимает Reset.
METHOD PRIVATE PositionLostLatchesFault
VAR
    fbTime   : FB_FakeTime;       // подменное время, старт 1 ч
    fbVlv    : FB_Valve;          // арматура под тестом
    stCmd    : ST_ValveCmd;       // команды HMI
    stRetain : ST_DeviceRetain;   // режим Manual по умолчанию, счётчики
    stCfg    : ST_ValveCfg;       // конфигурация (умолчания: Motorized, ZSO и ZSC)
    iStep    : INT;               // шаг цикла
END_VAR

(* ---- PositionLostLatchesFault.method.impl.st ---- *)
coUnit.TEST('Valve_PositionLost_LatchesFault');

fbVlv.xZso := TRUE;
// открыта
fbVlv(itfTime := fbTime, stCmd := stCmd, stRetain := stRetain, stCfg := stCfg);
fbVlv.xZso := FALSE;
// t0: провал ZSO
fbVlv(itfTime := fbTime, stCmd := stCmd, stRetain := stRetain, stCfg := stCfg);
FOR iStep := 1 TO 3 DO                                                  // t0 + 0,3 с
    fbTime.Advance(tStep := T#100MS);
    fbVlv(itfTime := fbTime, stCmd := stCmd, stRetain := stRetain, stCfg := stCfg);
END_FOR
fbVlv.xZso := TRUE;
fbTime.Advance(tStep := T#100MS);
// t0 + 0,4 с: вернулся
fbVlv(itfTime := fbTime, stCmd := stCmd, stRetain := stRetain, stCfg := stCfg);
AssertEquals_WORD(Expected := 0, Actual := fbVlv.stSts.stCommon.wFault, Message := 'short loss filtered');
AssertTrue(Condition := fbVlv.stSts.eState = E_ValveState.Open, Message := 'still Open');
fbVlv.xZso := FALSE;
fbTime.Advance(tStep := T#100MS);
// t1: ZSO пропал
fbVlv(itfTime := fbTime, stCmd := stCmd, stRetain := stRetain, stCfg := stCfg);
FOR iStep := 1 TO 4 DO                                                  // t1 + 0,4 с
    fbTime.Advance(tStep := T#100MS);
    fbVlv(itfTime := fbTime, stCmd := stCmd, stRetain := stRetain, stCfg := stCfg);
END_FOR
AssertEquals_WORD(Expected := 0, Actual := fbVlv.stSts.stCommon.wFault, Message := 'no fault before tLimitFilter');
AssertTrue(Condition := fbVlv.stSts.eState = E_ValveState.Open, Message := 'state held during the filter');
fbTime.Advance(tStep := T#100MS);
// t1 + 0,5 с
fbVlv(itfTime := fbTime, stCmd := stCmd, stRetain := stRetain, stCfg := stCfg);
AssertEquals_WORD(Expected := GVL_Const.VLV_FLT_POSITION_LOST, Actual := fbVlv.stSts.stCommon.wFault,
                  Message := 'PositionLost');
AssertTrue(Condition := fbVlv.stSts.eState = E_ValveState.Fault, Message := 'Fault state');
fbVlv.xZso := TRUE;
fbTime.Advance(tStep := T#100MS);
fbVlv(itfTime := fbTime, stCmd := stCmd, stRetain := stRetain, stCfg := stCfg);
AssertEquals_WORD(Expected := GVL_Const.VLV_FLT_POSITION_LOST, Actual := fbVlv.stSts.stCommon.wFault,
                  Message := 'latched after the limit switch returns');
stCmd.stCommon.xReset := TRUE;
fbVlv(itfTime := fbTime, stCmd := stCmd, stRetain := stRetain, stCfg := stCfg);
AssertEquals_WORD(Expected := 0, Actual := fbVlv.stSts.stCommon.wFault, Message := 'cleared by Reset');
AssertTrue(Condition := fbVlv.stSts.eState = E_ValveState.Open, Message := 'Open after Reset');

coUnit.TEST_FINISHED();

(* ---- PowerLossStopsWithoutFault.method.decl.st ---- *)
// Нет напряжения при открытии: Intermediate, выходы сняты, VLV_WRN_POWER_LOST, отказа нет; команда —
// RejectedInhibit; 12 с без напряжения (больше tTravel) отказа хода не дают. Напряжение вернулось:
// Manual стоит (цель снята); Auto снова ведёт к цели. Готовность для автоматики (Available,
// VLV_STS_AVAILABLE) в Auto есть только при напряжении.
METHOD PRIVATE PowerLossStopsWithoutFault
VAR
    fbTime   : FB_FakeTime;       // подменное время, старт 1 ч
    fbVlv    : FB_Valve;          // арматура под тестом
    stCmd    : ST_ValveCmd;       // команды HMI
    stRetain : ST_DeviceRetain;   // режим Manual по умолчанию, счётчики
    stCfg    : ST_ValveCfg;       // конфигурация (умолчания: Motorized, ZSO и ZSC)
    iStep    : INT;               // шаг цикла
END_VAR
